(* IEC 61131-3 sources: plcassist-cli/packages/volt-lsp-iec/test-corpus/awa-palletizer/Device/Plc Logic/Application/Library Manager/L_TS2P_TechModulesSynchronizingCamming (part 2) *)

(* ---- L_TS2P_FLYINGSAWSTATE.fb ---- *)
FUNCTION_BLOCK L_TS2P_FLYINGSAWSTATE EXTENDS L_TB2P_TechModuleBase
VAR_INPUT
	XUSEORIGINAL : BOOL;
	XENABLE : BOOL;
	XENABLEOPERATION : BOOL;
	XRESETERROR : BOOL;
	XQSPAPPLICATION : BOOL;
	XABORT : BOOL;
	XJOGPOS : BOOL;
	XJOGNEG : BOOL;
	XHOMEEXECUTE : BOOL;
	LROVERRIDE : LREAL := 1;
	SCCTRLBASICMOTION : L_TB2P_scCtrlBasicMotion;
	SCPAR : L_TS2P_scPar_FlyingSawState;
	SCACCESSPOINTS : L_TS2P_scAP_FlyingSawState;
	MASTERVALUES : L_MC1P_IAXIS_REF_MASTERVALUES;
	XSTARTFLYINGSAW : BOOL;
	XSYNCININSTANT : BOOL;
	XEXECUTENEXTCUT : BOOL;
	XEXECUTEGAP : BOOL;
	XSETCUTTINGLENGTHINSTANT : BOOL;
	LRCUTTINGLENGTH : LREAL;
	LRSYNCOVERRIDE : LREAL := 1;
	XSETMATERIALCOUNTER : BOOL;
	XMOVETOPARKPOS : BOOL;
	XRESUMETARGETPOS : BOOL;
	XRESETMARKSTACK : BOOL;
	SCTPRECDATA_MARKSENSOR : L_MC1P.L_MC1P_TpReceiveData;
END_VAR
VAR_OUTPUT
	XREADYFOROPERATION : BOOL;
	XOPERATIONENABLED : BOOL;
	XREADYFORMOTION : BOOL;
	XERROR : BOOL;
	XWARNING : BOOL;
	EERRORID : L_IE1P_Error;
	XSTOACTIVE : BOOL;
	XQSPACTIVE : BOOL;
	XABORTBUSY : BOOL;
	XABORTDONE : BOOL;
	XJOGGINGBUSY : BOOL;
	XHOMINGBUSY : BOOL;
	XHOMINGDONE : BOOL;
	XISHOMED : BOOL;
	ETMSTATE : L_TB2P_States := L_TB2P_States.DISABLED;
	SCSTATUSBASICMOTION : L_TB2P_scStatusBasicMotion;
	LRACTVEL : LREAL;
	LRSETVELOUT : LREAL;
	LRACTPOS : LREAL;
	LRSETPOSOUT : LREAL;
	LRACTFOLLOWINGERROR : LREAL;
	SCSIGNALFLOW : L_TS2P_scSF_FlyingSawState;
	XSYNCHRONISED : BOOL;
	XACCDECSYNC : BOOL;
	XINPOSITION : BOOL;
	XPOSITIONING : BOOL;
	LRMATERIALCOUNTER : LREAL;
	LRTARGETPOS : LREAL;
	LRCUTGAP : LREAL;
	LRACTIVECUTTINGLENGTH : LREAL;
	WMARKSINSTACK : WORD;
END_VAR
VAR_IN_OUT
	AXIS : AXIS_REF;
END_VAR
VAR
	XINTERNALCONTROLACTIVE_OLD : BOOL;
	XUSEORIGINAL_OLD : BOOL;
	ITFCONNECTORFLYINGSAW : L_TS2P_IConnectorFlyingSaw;
	TM_INT : L_TS2M_TM_FlyingSawState;
	SCPAR_INT : L_TS2P_scPar_FlyingSawState;
	_SCDATA_INT : L_TS2M_scData_FlyingSawState;
	_SCFMDATA_INT : L_TS2M_scData_FM_FlyingSaw;
	_UICALLMFUNIDXINPUT : UINT := 1;
	_UICALLMFUNIDXOUTPUT : UINT := 1;
	_MCCALL : L_UM1P_MCCall;
	_ASCINPUT : ARRAY [1.._MCCall.c_BufferDepthInput] OF L_TS2P_FlyingSawStateIn;
	_ASCOUTPUT : ARRAY [1.._MCCall.c_BufferDepthOutput] OF L_TS2P_FlyingSawStateOut;
	_ASCPARCORE : ARRAY [1.._MCCall.c_BufferDepthInput] OF L_TS2P_scPar_FlyingSawState;
	_ASCACCESSPOINTSCORE : ARRAY [1.._MCCall.c_BufferDepthInput] OF L_TS2P_scAP_FlyingSawState;
	_ASCSIGNALFLOWCORE : ARRAY [1.._MCCall.c_BufferDepthOutput] OF L_TS2P_scSF_FlyingSawState;
	_ASCDATACORE : ARRAY [1.._MCCall.c_BufferDepthInput] OF L_TS2M_scData_FlyingSawState;
	_ASCDATAFMCORE : ARRAY [1.._MCCall.c_BufferDepthInput] OF L_TS2M_scData_FM_FlyingSaw;
	_SCINPUTVISU : L_TS2P_FlyingSawStateIn;
	_PSCINPUTVISU : POINTER TO L_TS2P_FlyingSawStateIn := ADR(_scInputVisu);
	_PSCOUTPUTVISU : POINTER TO L_TS2P_FlyingSawStateOut := ADR(_ascOutput[1]);
	_PSCPARVISU : POINTER TO L_TS2P_scPar_FlyingSawState := ADR(scPar_int);
	_PSCDATAVISU : POINTER TO L_TS2M_scData_FlyingSawState := ADR(_scData_int);
	_PSCFMDATAVISU : POINTER TO L_TS2M_scData_FM_FlyingSaw := ADR(_scFMData_int);
	_PSCFMSFVISU : POINTER TO L_TS2P_scSF_FlyingSawState;
	ITFBASICMOTIONBASE : L_TB2P.L_TB2P_IBasicMotionBase;
	ITFFLYINGSAWPROCESSINGEXTENSION : L_TS2P_IFlyingSawProcessing;
	ITFITECHMODULEINTERNAL : L_TB2P_ITechModuleInternal;
	LRJERKDEC : LREAL;
	LRJOGGINGJERKDEC : LREAL;
	REMAININGTIMEOFPROFILE : LREAL;
	REMAININGTIMEOFPROFILEAVAILABLE : BOOL;
END_VAR
END_FUNCTION_BLOCK

METHOD CALL_ABC
VAR_INPUT
	ITFTECHMODULE : L_TB2P.L_TB2P_IBasicMotionBase;
	XQSPAPPLICATION : BOOL;
	XHALT : BOOL;
	XABORT : BOOL;
	XHOMEEXECUTE : BOOL;
	XJOGPOS : BOOL;
	XJOGNEG : BOOL;
	XFINISHPOSITIONING : BOOL;
	XMOVEVELEXECUTE : BOOL;
	XMOVEABSEXECUTE : BOOL;
	XMOVERELEXECUTE : BOOL;
	XENABLEOPERATION : BOOL;
	XRESETERROR : BOOL;
	XENABLEPOSITIVE : BOOL;
	XENABLENEGATIVE : BOOL;
	XDISABLESWLIMIT : BOOL;
	LROVERRIDE : LREAL;
	LROVERRIDEACC : LREAL;
	LROVERRIDEJERK : LREAL;
	XRESETHOMEPOSITION : BOOL;
	XCONTINUOUSUPDATE : BOOL;
	LRPOS_DIST : LREAL;
	LRVEL : LREAL;
	LRACC : LREAL;
	LRDEC : LREAL;
	LRJERK : LREAL;
	EDIRECTION : L_TB2P.MC_DIRECTION;
	SCHOMEEXTTP : L_TB2P.MC_TRIGGER_REF;
	XHOMEABSSWITCH : BOOL;
	XSPECIALABORTBEHAVIOR : BOOL;
	LRABORTDEC : LREAL;
	LRABORTJERK : LREAL;
END_VAR
VAR_OUTPUT
	XERROR : BOOL;
	EERRORID : L_TB2P.L_IE1P_Error;
	XFUNBUSY : BOOL;
	XFUNDONE : BOOL;
	XFUNCOMMANDABORTED : BOOL;
	EFUNSTATEACT : L_TB2P.L_MC1P_ABC_State;
	ECONTROLMODE : L_TB2P.L_MC1P_ControlMode;
	XISHOMED : BOOL;
	XHWLIMITSWITCHNEG : BOOL;
	XHWLIMITSWITCHPOS : BOOL;
	XSWLIMITENABLED : BOOL;
	XSWLIMITSWITCHNEG : BOOL;
	XSWLIMITSWITCHPOS : BOOL;
	EAXISTYPE : L_TB2P.L_MC1P_DriveType;
	EAXISSTATE : L_TB2P.L_MC1P_AXIS_STATE;
	XSTOACTIVE : BOOL;
	XREADYFOROPERATION : BOOL;
	XOPERATIONENABLED : BOOL;
	XREADYFORMOTION : BOOL;
	XAXISWARNING : BOOL;
	XAXISERROR : BOOL;
	EAXISERRORID : L_TB2P.L_IE1P_Error;
	XDRIVEWARNING : BOOL;
	XDRIVEERROR : BOOL;
	DWDRIVEERRORID : DWORD;
	LRACTPOS : LREAL;
	LRACTVEL : LREAL;
	LRSETPOSOUT : LREAL;
	LRSETVELOUT : LREAL;
	LRACTFOLLOWINGERROR : LREAL;
	XINPOSITION : BOOL;
	XSTANDSTILLSETVELOCITY : BOOL;
	XSTANDSTILLACTVELOCITY : BOOL;
	XCONSTANTVELOCITY : BOOL;
	XACCELERATING : BOOL;
	XDECELERATING : BOOL;
	XDIRECTIONPOSITIVE : BOOL;
	XDIRECTIONNEGATIVE : BOOL;
	XAXISAVAILABLE : BOOL;
END_VAR
VAR_IN_OUT
	AXIS : AXIS_REF;
END_VAR
END_METHOD

METHOD GET_PAP : POINTER TO L_TB2P_scAP_TM_MotionControl
END_METHOD

METHOD GET_PDATA : POINTER TO L_TS2M_scData_FlyingSawState
END_METHOD

METHOD GET_PFMDATA : POINTER TO L_TS2M_scData_FM_FlyingSaw
END_METHOD

METHOD GET_PPAR : POINTER TO L_TB2P_scPar_TM_MotionControl
END_METHOD

METHOD GET_PSF : POINTER TO L_TB2P_scSF_TM_MotionControl
END_METHOD

METHOD CLUTCH
VAR_INPUT
	ITFTECHMODULE : L_TS2P_IFlyingSawProcessing;
	XENABLE : BOOL;
	XSYNCVEL : BOOL := FALSE;
	XSYNCPOS : BOOL;
	XSYNCOUTINSTANT : BOOL;
	LRSYNCVEL : LREAL := 10;
	LRSYNCACC : LREAL := 100;
	LRSYNCDEC : LREAL := 100;
	LRSYNCJERK : LREAL := 10000;
	LRCYCMASTERPOS : LREAL;
	LRCYCMASTERVEL : LREAL;
	LRCYCMASTERACC : LREAL;
	LRSETSLAVEPOS : LREAL;
	LRSETSLAVEVEL : LREAL;
	LRSETSLAVEACC : LREAL;
END_VAR
VAR_OUTPUT
	EERRORID : L_IE1P.L_IE1P_Error;
	XERROR : BOOL;
	XBUSY : BOOL;
	XDONE : BOOL;
	XACCDECSYNC : BOOL;
	XVELSYNCHRONISED : BOOL;
	XPOSSYNCHRONISED : BOOL;
	LRSETSLAVEPOSOUT : LREAL;
	LRSETSLAVEVELOUT : LREAL;
	LRSETSLAVEACCOUT : LREAL;
	XPROFILERESETTIMEVALID : BOOL;
	LRPROFILERESETTIME : LREAL;
END_VAR
END_METHOD

METHOD EXECUTEGAP
VAR_INPUT
	ITFTECHMODULE : L_TS2P_IFlyingSawProcessing;
	XENABLE : BOOL;
	LRSYNCVEL : LREAL := 10;
	LRSYNCACC : LREAL := 100;
	LRSYNCDEC : LREAL := 100;
	LRSYNCJERK : LREAL := 10000;
	XEXECUTEGAP : BOOL;
	XAUXEXECUTEGAP : BOOL := FALSE;
	LRCYCMASTERPOS : LREAL;
	LRCYCMASTERVEL : LREAL;
	LRCYCMASTERACC : LREAL;
	LRSETSLAVEPOS : LREAL;
	LRSETSLAVEVEL : LREAL;
	LRSETSLAVEACC : LREAL;
END_VAR
VAR_OUTPUT
	EERRORID : L_IE1P.L_IE1P_Error;
	XERROR : BOOL;
	XBUSY : BOOL;
	XDONE : BOOL;
	XACCDECSYNC : BOOL;
	XVELSYNCHRONISED : BOOL;
	XPOSSYNCHRONISED : BOOL;
	LRSETSLAVEPOSOUT : LREAL;
	LRSETSLAVEVELOUT : LREAL;
	LRSETSLAVEACCOUT : LREAL;
	XPROFILERESETTIMEVALID : BOOL;
	LRPROFILERESETTIME : LREAL;
END_VAR
END_METHOD

METHOD MARKSTACK_GETMARK
VAR_INPUT
	ITFTECHMODULE : L_TS2P_IFlyingSawProcessing;
	XENABLE : BOOL;
	XGETMARK : BOOL;
	XRESETGETMARK : BOOL;
	XRESETMARKSTACK : BOOL;
	LRCYCSETPOS : LREAL;
	LRCYCSETVEL : LREAL;
END_VAR
VAR_OUTPUT
	XMARKSTACKFULL : BOOL;
	XMARKSTACKEMPTY : BOOL;
	WMARKSINSTACK : WORD;
	XMARKVALID : BOOL;
	LRMARKPOSOUT : LREAL;
END_VAR
END_METHOD

METHOD MARKSTACK_SETMARK
VAR_INPUT
	ITFTECHMODULE : L_TS2P_IFlyingSawProcessing;
	XENABLE : BOOL;
	XSETMARK : BOOL;
	LRMARKPOS : LREAL;
	XRESETMARKSTACK : BOOL;
	LRCYCSETPOS : LREAL;
	LRCYCSETVEL : LREAL;
END_VAR
VAR_OUTPUT
	XMARKSTACKFULL : BOOL;
	XMARKSTACKEMPTY : BOOL;
	WMARKSINSTACK : WORD;
	XNEWMARKRECEIVED : BOOL;
END_VAR
END_METHOD

METHOD POSITIONING
VAR_INPUT
	ITFTECHMODULE : L_TS2P_IFlyingSawProcessing;
	XENABLE : BOOL;
	XMOVETOTARGETPOS : BOOL;
	LRTARGETPOS : LREAL;
	LRPOSITIONINGVEL : LREAL;
	LRPOSITIONINGACC : LREAL;
	LRPOSITIONINGDEC : LREAL;
	LRPOSITIONINGJERK : LREAL;
	LRSETSLAVEPOS : LREAL;
	LRSETSLAVEVEL : LREAL;
	LRSETSLAVEACC : LREAL;
	LRCORRECTTIMEBASE : LREAL := 0;
	LROVERRIDE : LREAL := 1.0;
END_VAR
VAR_OUTPUT
	EERRORID : L_IE1P.L_IE1P_Error;
	XERROR : BOOL;
	XBUSY : BOOL;
	XDONE : BOOL;
	XPOSITIONING : BOOL;
	XINPOSITION : BOOL;
	LRSETSLAVEPOSOUT : LREAL;
	LRSETSLAVEVELOUT : LREAL;
	LRSETSLAVEACCOUT : LREAL;
	XPROFILERESETTIMEVALID : BOOL;
	LRPROFILERESETTIME : LREAL;
END_VAR
END_METHOD

METHOD REQUESTINTERFACE : BOOL
VAR_INPUT
	ID : DINT;
	PITFUNKNOWN : POINTER TO L_UBUP.L_UBUP_IUnknown;
END_VAR
END_METHOD

METHOD CALLFUNCTION
VAR_INPUT
	UIINPUTDATAIDX : UINT;
	UIOUTPUTDATAIDX : UINT;
END_VAR
END_METHOD

METHOD COPYINPUTS : BOOL
VAR_INPUT
	IDX : WORD;
END_VAR
END_METHOD

METHOD COPYOUTPUTS : BOOL
VAR_INPUT
	IDX : WORD;
END_VAR
END_METHOD

METHOD FUNCTIONWASCALLEDTWICE : BOOL
VAR_INPUT
	IDX : WORD;
END_VAR
END_METHOD

METHOD HANDLESTANDARDCALL : BOOL
END_METHOD

METHOD SYNCOUTPUTS
VAR_INPUT
	UICOPYOUTPUTFROMIDX : UINT;
	UICOPYOUTPUTTOIDX : UINT;
END_VAR
END_METHOD

METHOD FB_INIT : BOOL
VAR_INPUT
	BINITRETAINS : BOOL;
	BINCOPYCODE : BOOL;
END_VAR
END_METHOD

METHOD CALL_INTERNALCTRL
END_METHOD

(* ---- L_TS2P_INVERTGEARFACTOR.fb ---- *)
FUNCTION_BLOCK L_TS2P_INVERTGEARFACTOR
VAR_INPUT
	XINVERTGEARFACTOR : BOOL;
	LRCYCLELENGTHX : LREAL := 1.0;
	LRCYCLELENGTHY : LREAL := 1.0;
	LRCOUPLINGX : LREAL := 1.0;
	LRCOUPLINGY : LREAL := 1.0;
	XDISABLETOLERANCEINVERTGEARFACTOR : BOOL;
	LRTOLERANCEINVERTGEARFACTOR : LREAL := 0;
END_VAR
VAR_OUTPUT
	XINVERTGEARFACTORACTIVE : BOOL;
	LRCYCLELENGTHX_OUT : LREAL;
	LRCYCLELENGTHY_OUT : LREAL;
	LRCOUPLINGX_OUT : LREAL;
	LRCOUPLINGY_OUT : LREAL;
	XWARNING : BOOL;
	EERRORID : L_IE1P_Error;
END_VAR
VAR_IN_OUT
	AXIS : AXIS_REF;
END_VAR
VAR
	XINWINDOW : BOOL;
END_VAR
END_FUNCTION_BLOCK

(* ---- L_TS2P_MARKQUEUE.fb ---- *)
FUNCTION_BLOCK L_TS2P_MARKQUEUE
VAR_INPUT
	XENABLE : BOOL;
	XLOADMARKPOS : BOOL;
	LRMARKPOS : LREAL;
	XGETNEXTMARK : BOOL;
	XRESETGETNEXTMARK : BOOL;
	XRESETMARKQUEUE : BOOL;
	LRCYCSETPOS : LREAL;
	LRCYCSETVEL : LREAL;
END_VAR
VAR_OUTPUT
	XQUEUEISFULL : BOOL;
	XQUEUEISEMPTY : BOOL;
	XNEWMARKRECEIVED : BOOL;
	WMARKSINQUEUE : WORD;
	XMARKVALID : BOOL;
	LRMARKPOSOUT : LREAL;
END_VAR
VAR
	FB_MB1P_STACK : L_MB1P_Stack;
	XTRACKMARK : BOOL;
	XENABLE_OLD : BOOL;
	XRESETMARKQUEUE_OLD : BOOL;
	XGETNEXTMARK_OLD : BOOL;
	XRESETGETNEXTMARK_OLD : BOOL;
	C_LRMATERIALCOUNTERCYCLELENGTH : LREAL := (16#4FFFFFFFFFFFFFFF * 1E-08);
END_VAR
END_FUNCTION_BLOCK

(* ---- L_TS2P_MARKSTACK.fb ---- *)
FUNCTION_BLOCK L_TS2P_MARKSTACK
VAR_INPUT
	XENABLE : BOOL;
	TPRECDATAIN : L_MC1P_TpReceiveData;
	LRACTVELMATERIAL : LREAL;
	LRACTPOSITIONTPAXIS : LREAL;
	LRCYCLELENGTHTPAXIS : LREAL;
	LRMARKSTACKLENGTH : LREAL;
	LRTASKCYCLE : LREAL;
END_VAR
VAR_OUTPUT
	TPRECDATAOUT : L_MC1P_TpReceiveData;
	XERROR : BOOL := FALSE;
	EERRORID : WORD;
	LRTPDIFFOUT : LREAL;
END_VAR
VAR
	ALRINTEGRATORSTARTPOS : ARRAY [1..64] OF LREAL := [64(0)];
	ALRLASTSCAN : ARRAY [1..64] OF LREAL := [64(0)];
	ALRDUMMY : ARRAY [1..64] OF LREAL := [64(0)];
	AXTPVALID : ARRAY [1..64] OF BOOL := [64(FALSE)];
	AXDUMMY : ARRAY [1..64] OF BOOL := [64(FALSE)];
	ADWACTTIMESTAMP : ARRAY [1..64] OF DWORD := [64(0)];
	ADWRECTIMESTAMP : ARRAY [1..64] OF DWORD := [64(0)];
	ADWDUMMY : ARRAY [1..64] OF DWORD := [64(0)];
	XREGISTERFULL : BOOL := FALSE;
	XINIT : BOOL := TRUE;
	WCOUNTER : WORD;
	WCOUNTERIN : WORD := 1;
	WCOUNTEROUT : WORD := 1;
	LRINTEGRATORPOS : LREAL := 0;
	LRCYCPOSDIFF : LREAL := 0;
	LRPOSTOREGISTEREND : LREAL := 0;
	XTPRECEIVEDINOLD : BOOL;
	LRMARKSTACKLENGTHOLD : LREAL;
	LRACTPOSITIONTPAXISCOMP : LREAL;
	LRACTTPPOSITIONOUT_INT : LREAL;
	DWDEADTIMESTACKOUT : DWORD;
	LRINTEGRATORLENGTH : LREAL := 10000000000.0;
END_VAR
END_FUNCTION_BLOCK

METHOD CALL_INITMARKSTACK
END_METHOD

(* ---- L_TS2P_MARKSTACKFLYINGSAW.fb ---- *)
FUNCTION_BLOCK L_TS2P_MARKSTACKFLYINGSAW
VAR
	FB_MB1P_STACK : L_MB1P_Stack_FlyingSaw;
	XTRACKMARK : BOOL;
	XMARKVALID_INT : BOOL;
	XENABLE_OLD : BOOL;
	XRESETMARKSTACK_OLD : BOOL;
	XGETMARK_OLD : BOOL;
	XSETMARK_OLD : BOOL;
	XRESETGETMARK_OLD : BOOL;
	C_LRMATERIALCOUNTERCYCLELENGTH : LREAL := (16#4FFFFFFFFFFFFFFF * 1E-08);
END_VAR
END_FUNCTION_BLOCK

METHOD DISABLE
END_METHOD

METHOD RESETMARKSTACK
END_METHOD

METHOD GETMARK
VAR_INPUT
	XENABLE : BOOL;
	XGETMARK : BOOL;
	XRESETGETMARK : BOOL;
	XRESETMARKSTACK : BOOL;
	LRCYCSETPOS : LREAL;
	LRCYCSETVEL : LREAL;
END_VAR
VAR_OUTPUT
	XMARKSTACKFULL : BOOL;
	XMARKSTACKEMPTY : BOOL;
	WMARKSINSTACK : WORD;
	XMARKVALID : BOOL;
	LRMARKPOSOUT : LREAL;
END_VAR
END_METHOD

METHOD SETMARK
VAR_INPUT
	XENABLE : BOOL;
	XSETMARK : BOOL;
	LRMARKPOS : LREAL;
	XRESETMARKSTACK : BOOL;
	LRCYCSETPOS : LREAL;
	LRCYCSETVEL : LREAL;
END_VAR
VAR_OUTPUT
	XMARKSTACKFULL : BOOL;
	XMARKSTACKEMPTY : BOOL;
	WMARKSINSTACK : WORD;
	XNEWMARKRECEIVED : BOOL;
END_VAR
END_METHOD

(* ---- L_TS2P_MARKWINDOWRELATIVE.fb ---- *)
FUNCTION_BLOCK L_TS2P_MARKWINDOWRELATIVE
VAR_INPUT
	XENABLE : BOOL;
	LRTPWINDOWSIZE : LREAL;
	LRSETOFFSETTPWINDOW : LREAL;
	LRCYCVEL : LREAL;
	TPRECDATAIN : L_MC1P_TpReceiveData;
	LRSTARTPOSITION : LREAL;
	LRCYCLELENGTH : LREAL;
	XTEACHMARKWINDOW : BOOL;
	DWMAXTPNOTDETECTED : DWORD;
	LRTASKCYCLE : LREAL;
END_VAR
VAR_OUTPUT
	TPRECDATAOUT : L_MC1P_TpReceiveData;
	XTPWINDOWOPEN : BOOL;
	XTPWINDOWOPENCOMP : BOOL;
	LRTPDELTAPOSCOMP : LREAL;
	XTPINWINDOW : BOOL;
	XTPNOTINWINDOW : BOOL;
	XTPNOTDETECTED : BOOL;
	XTPSENSORTEACHED : BOOL;
	XMAXTPNOTDETECTED : BOOL;
END_VAR
VAR
	LRMARKWINDOWINTEGRATOROLD : LREAL;
	XTPNOTDETECTEDINTERNAL : BOOL;
	LRLOWERWINDOW : LREAL;
	LRUPPERWINDOW : LREAL;
	XTEACHTPSENSOROLD : BOOL;
	DWMISSEDTPCOUNTER : DWORD;
	XTPISINWINDOW : BOOL;
	LRDEADTIMEPOSDIFF : LREAL;
	LRUPPERWINDOWCOMP : LREAL;
	XTPCOMPWINDOWOPEN : BOOL;
	XTPCOMPWINDOWOPENOLD : BOOL := FALSE;
	LRLOWERWINDOWCOMP : LREAL;
	XTPRECEIVEDOLD : BOOL;
	XTPRECEIVEDINTERNAL : BOOL;
	LRTPWINDOWSIZE_INT : LREAL;
	LRMARKWINDOWINTEGRATOR : LREAL := 0;
	LRDEADTIMETP : LREAL;
	LRACTUALTPPOSITION : LREAL;
END_VAR
END_FUNCTION_BLOCK

(* ---- L_TS2P_MASTERVALUECORRECTION.fb ---- *)
FUNCTION_BLOCK L_TS2P_MASTERVALUECORRECTION
VAR_INPUT
	XAXIS : POINTER TO L_MC1P_IAXIS_REF_MASTERVALUES;
	XENABLE : BOOL;
	XENABLECORRECTION : BOOL;
	XRESETERROR : BOOL;
	LRSETVELIN : LREAL;
	LRACTPOSITIONTOOL : LREAL;
	LRCYCLELENGTHTOOL : LREAL;
	TPRECDATA : L_MC1P_TpReceiveData;
	XLOADREGPOS : BOOL;
	LRLOADREGPOS : LREAL;
	LRSENSORTOOLDIST : LREAL;
	LRMARKDIST : LREAL;
	LRMAXCORRNEG : LREAL;
	LRMAXCORRPOS : LREAL;
	ESOURCEFORCORRWINDOW : L_TS2P_SourceForCorrWindow;
	LRUPPERCORRPOS : LREAL;
	LRLOWERCORRPOS : LREAL;
	DWGEARINGNUMERATORY : DWORD := 1;
	DWGEARINGDENOMINATORY : DWORD := 1;
	XSYNCHRONISED : BOOL;
	LRACTOFFSETMASTERIN : LREAL;
	LRACTOFFSETSLAVEIN : LREAL;
	XTEACHMARKWINDOW : BOOL;
	XENABLEMARKWINDOW : BOOL;
	LRMARKWINDOWSIZE : LREAL;
	LRSETOFFSETMARKWINDOW : LREAL;
	DWMAXNUMBERVIRTUALMARKS : DWORD;
	LRGEARFACTORCORRGAIN : LREAL;
	LRMAXGEARFACTORCORR : LREAL;
	XGEARFACTORCORR : BOOL;
	XGEARFACTORCORRHOLD : BOOL;
	XENABLETOOLCORRECTION : BOOL;
	LRTRANSMITCYCLESSETPOS : LREAL;
	DIDEADTIMECOMP : DINT;
	LRCORRVEL : LREAL;
	LRCORRACC : LREAL;
	LRCORRDEC : LREAL;
	LRCORRJERK : LREAL;
	ECORRMODE : L_TS2P_CorrectionMode;
	ECORRMODEOLD : L_TS2P_CorrectionMode;
END_VAR
VAR_OUTPUT
	CORRECTEDXAXIS : L_MC1P_IAXIS_REF_MASTERVALUES;
	LRACTVEL : LREAL;
	XERROR : BOOL;
	XWARNING : BOOL;
	EERRORID : WORD;
	XCORRLIMITED : BOOL;
	LRACTMARKERROR : LREAL;
	LRACTMARKDIST : LREAL;
	XINITDONE : BOOL;
	XCORRACTIVE : BOOL;
	XMARKRECEIVED : BOOL;
	LRSENSORACTPOS : LREAL;
	LRSENSORSETPOS : LREAL;
	XMARKWINDOWOPEN : BOOL;
	XMARKOUTOFWINDOW : BOOL;
	XMARKNOTDETECTED : BOOL;
	XMARKWINDOWTEACHED : BOOL;
	LRGEARFACTORCORR : LREAL;
	XGEARFACTORCORRLIMITED : BOOL;
	XCORRNEXTCYCLE : BOOL;
END_VAR
VAR_IN_OUT
	YAXIS : AXIS_REF;
END_VAR
VAR
	FB_L_TB2P_TP_CONVERTER : L_TB2P_TP_Converter;
	FB_L_TS2P_MARKWINDOWRELATIVE : L_TS2P_MarkWindowRelative;
	FB_L_TS2P_TPVIRTUALACTPOS : L_TS2P_TpVirtualActPos;
	FB_L_TS2P_MARKSTACK : L_TS2P_MarkStack;
	FB_L_MC1P_TPCALCDIFF : L_MC1P_TpCalcDiff;
	FB_L_TS2P_TPLIMITDIFF : L_TS2P_TpLimitDiff;
	FB_L_TS2P_DISTCORRECTIONWINDOW : L_TS2P_DistCorrectionWindow;
	FB_L_MC1P_SETAXISREFMASTERVALUES : L_MC1P_SetAxisRefMasterValues;
	FB_PROFILEGENERATOR : L_MC1P_ProfileGenerator;
	FB_INTEGRATOR : L_MC1P_IntegrateAxis;
	SCPROFILEPARAMETER : L_MC1P_ProfileParameter;
	FB_RAMPGENERATORGEARFACTOR : L_MC1P_RampGenerator;
	LRSENSORSETPOS_INT : LREAL;
	LRGEARINGFAKTOR : LREAL := 1.0;
	LRTPDIFFERENCE_INT : LREAL;
	XTPINWINDOW : BOOL;
	XVALUESTOREDTPCONVERTER : BOOL;
	XVALUESTOREDTPCONVERTEROLD : BOOL;
	XVALUESTOREDMARKWINDOW : BOOL;
	XVALUESTOREDMISSEDMARKS : BOOL;
	XVALUESTOREDMARKSTACK : BOOL;
	XVALUESTOREDCALCDIFF : BOOL;
	XVALUESTOREDLIMIT : BOOL;
	LRCORRRESIDUAL : LREAL;
	LRTPACTPOSITION_INT : LREAL;
	LRTPDIFFERENCELIM_INT : LREAL;
	LROFFSETPOSCTRL_INT : LREAL;
	LRCYCVELIN_INT : LREAL;
	LRSETCORRECTEDPOSOUT_INT : LREAL;
	LRMASTERSETPOSOLD_INT : LREAL;
	LRCORRPOSOUTOLD_INT : LREAL;
	LRVELOUT_INT : LREAL;
	XCORRACTIVE_INT : BOOL;
	XINIT : BOOL := TRUE;
	XTPCORRECTIONACTIVE : BOOL := FALSE;
	LRTPAXISSETPOS : LREAL;
	LRMARKDIST_INT : LREAL;
	XZERO : BOOL;
	XHOMINGDONE : BOOL;
	XSTARTREFERENCEACTIVE : BOOL;
	XHOMINGACTIVE : BOOL := FALSE;
	XMARKDISTCHANGED : BOOL;
	XENABLE_OLD : BOOL;
	XTPRECEIVEDOUT_INTOLD : BOOL;
	XSTARTFIRSTCORRECTION : BOOL;
	LRTPDIFFERENCELIM2_INT : LREAL;
	XCORRECTIONBUSYOLD : BOOL;
	LRTPACTPOSIN_OLD : LREAL;
	LRTPSETPOSIN_OLD : LREAL;
	LRTPAXISACTPOS_OLD : LREAL;
	LRCYCLELENGTH : LREAL;
	ICOUNTER : INT := 0;
	LRSETPOSITIONOLD : LREAL;
	LRCYCLELENGTHTP : LREAL;
	LRTPACTPOSITIONOLD : LREAL;
	XFIRSTTOUCHPROBE : BOOL := TRUE;
	LRSENSORTOOLDISTANCE_INT : LREAL;
	LRMARKSTACKLENGTH : LREAL;
	LRTPDIFFERENCELIMITOUT_INT : LREAL;
	XTPNOTDETECTED_INT : BOOL;
	XMAXTPNOTDETECTED : BOOL;
	LRGEARINGFAKTOROLD : LREAL;
	LRGEARFACTORINTEGRATOR : LREAL;
	LRGEARFACTORGAIN : LREAL := 1;
	LRGEARFACTORNUMERATORCORR : LREAL;
	LRGEARFACTORNUMERATORCORRLIMITED : LREAL;
	LRGEARFACTORDENOMINATOR : LREAL;
	LRGEARFACTORNUMERATOR : LREAL;
	LRTOTALSTACKDIFFERENCEOUT_INT : LREAL := 0;
	LCORRECTIONVELIN : LREAL;
	LRSETPOSCORROUT_OLD : LREAL;
	LRDELTAGEARFACTORCORR : LREAL;
	XTPSENSORTEACHEDOLD : BOOL;
	XTPSENSORTEACHEDATLASTMARK : BOOL;
	XCALCMARKDISTINITIALISED : BOOL;
	XTEACHTPSENSOROLD : BOOL;
	LRTPDEADTIMEDIFF : LREAL;
	XTPRECEIVEDOUTOLD_INT : BOOL;
	LRMARKDISTINTEGRATOR : LREAL;
	LRTPAXISCOMPFACTOR : LREAL;
	LRTPAXISDELAYCYCLE : LREAL;
	XENABLEOLD : BOOL;
	XTPRECEIVEDINOLD_INT : BOOL;
	TPRECDATAMARKWINDOW : L_MC1P_TpReceiveData;
	TPRECDATAMARKSTACK : L_MC1P_TpReceiveData;
	LRMASTERACTPOSITIONOLD_INT : LREAL;
	XFIRSTVALUESTORED : BOOL := FALSE;
	LRSETINTEGRATEDPOSITIONOLD : LREAL;
	XRESETERROROLD : BOOL;
	LRTPDIFF : LREAL;
	LRVELDIFF : LREAL;
	LRVELCOMP : LREAL;
	SETPOSITIONFORSYNCOLD : LREAL;
	LRMARKDISTOLD : LREAL;
END_VAR
END_FUNCTION_BLOCK

METHOD CALL_CALCACTMARKDIST
END_METHOD

METHOD CALL_CALCMARKERROR
END_METHOD

METHOD CALL_CORRECTIONPOS
END_METHOD

METHOD CALL_CORRECTIONPROFILE
END_METHOD

METHOD CALL_ENABLEREGISTERCONTROL
END_METHOD

METHOD CALL_ERRORHANDLER
END_METHOD

METHOD CALL_FB
VAR_IN_OUT
	YAXIS : AXIS_REF;
END_VAR
END_METHOD

METHOD CALL_GEARFACTORCORRECTION
END_METHOD

METHOD CALL_GEARING
END_METHOD

METHOD CALL_INPUT
END_METHOD

METHOD CALL_LIMIT
END_METHOD

METHOD CALL_MARKDISTCHANGE
END_METHOD

METHOD CALL_MARKSENSORPOS
END_METHOD

METHOD CALL_MARKSTACK
END_METHOD

METHOD CALL_MARKWINDOW
VAR_IN_OUT
	YAXIS : AXIS_REF;
END_VAR
END_METHOD

METHOD CALL_NOTENABLE
END_METHOD

METHOD CALL_OUTPUT
END_METHOD

METHOD CALL_RESET
END_METHOD

METHOD CALL_RESETOUTPUTS
END_METHOD

METHOD CALL_SETAXISREFMASTERVALUES
END_METHOD

METHOD CALL_TPCONVERTER
END_METHOD

METHOD CALL_VIRTUALACTPOS
END_METHOD

METHOD GET_ACTMARKERRORLIMITED : LREAL
END_METHOD

METHOD GET_ACTUALMARKDIST : LREAL
END_METHOD

METHOD GET_CORRREGPOS : LREAL
END_METHOD

METHOD GET_INTEGRATORREGPOS : LREAL
END_METHOD

METHOD GET_MARKERRORUNLIMITED : LREAL
END_METHOD

METHOD GET_MARKPOSITIONINREGISTER : LREAL
END_METHOD

METHOD GET_MARKRECEIVEUNLIMITED : BOOL
END_METHOD

METHOD GET_MARKRECEIVEDLIMITED : BOOL
END_METHOD

METHOD GET_MARKWINDOWCOMP : BOOL
END_METHOD

METHOD GET_REGISTERINPUTVEL : LREAL
END_METHOD

METHOD GET_SETVELOCITYREGISTER : LREAL
END_METHOD

METHOD GET_LRMARKSTACKLENGTH : LREAL
END_METHOD

METHOD SETTPCOMPFACTOR : LREAL
END_METHOD

METHOD SETTPDELAYCYCLE : LREAL
END_METHOD

(* ---- L_TS2P_MATERIALCOUNTER.fb ---- *)
FUNCTION_BLOCK L_TS2P_MATERIALCOUNTER
VAR_INPUT
	XENABLE : BOOL;
	LRPOSIN : LREAL;
	LRTASKCYCLE : LREAL;
	LRPOSINSLAVE : LREAL;
	LRCYCLELEN : LREAL;
	XLOADSTARTPOS : BOOL;
	XSETMATERIALCOUNTER : BOOL;
	LRSETMATERIALPOS : LREAL;
	XLOADDELTAPOS : BOOL;
	LRSETDELTAPOS : LREAL;
	XSTARTFLYINGSAW : BOOL;
END_VAR
VAR_OUTPUT
	LNMATERIALPOS_E8 : LINT;
	LRMATERIALCOUNTER : LREAL;
	LRDELTAMATERIALPOS : LREAL;
END_VAR
VAR_IN_OUT
	AXIS : AXIS_REF;
END_VAR
VAR
	LNMODULOPOS_E8 : LINT;
	LNMODULOPOSOLD_E8 : LINT;
	LNCYCLELEN_E8 : LINT;
	LNPOSXDIFF : LINT;
	LNMATERIALPOS_E8_OLD : LINT;
	LNDELTAMATERIALPOS : LINT;
	XSETMATERIALCOUNTER_OLD : BOOL;
	XENABLE_OLD : BOOL;
END_VAR
END_FUNCTION_BLOCK

(* ---- L_TS2P_MULTICAMSEQUENCER.fb ---- *)
FUNCTION_BLOCK L_TS2P_MULTICAMSEQUENCER
VAR_INPUT
	XENABLE : BOOL;
	XCAMSEQUENCER : BOOL;
	EMODE : L_TS2P_CamSequenceMode;
	XCAMCHANGEINSTANT : BOOL;
	XLOADCAMTABLE : BOOL;
	WSETCAMTABLE : WORD;
	XENDOFPROFILEIN : BOOL;
	CAMTABLE1 : MC_CAM_REF;
	CAMTABLE2 : MC_CAM_REF;
	CAMTABLE3 : MC_CAM_REF;
	CAMTABLE4 : MC_CAM_REF;
END_VAR
VAR_OUTPUT
	XDONE : BOOL;
	XBUSY : BOOL;
	XERROR : BOOL;
	EERRORID : L_IE1P_Error;
	WACTIVECAMTABLE : WORD;
	CAMTABLEOUT : MC_CAM_REF;
	XCAMTABLEVALID : BOOL;
END_VAR
VAR
	WFMSTATE : WORD := 0;
	XINITSTATE : BOOL;
	XENABLE_OLD : BOOL;
	XLOADCAMTABLE_OLD : BOOL;
	XENDOFPROFILEIN_OLD : BOOL;
	XCAMSEQUENCER_OLD : BOOL;
	XCAMCHANGEINSTANT_OLD : BOOL;
	XCAMSEQUENCERACTIVE : BOOL;
END_VAR
END_FUNCTION_BLOCK

METHOD CALL_ERRORHANDLER
END_METHOD

METHOD CALL_FBMETHODS
END_METHOD

METHOD CALL_OUTPUT
END_METHOD

METHOD CALL_RESETCOMMANDS
END_METHOD

METHOD CALL_RESETOUTPUT
END_METHOD

METHOD CALL_STATEMACHINE
END_METHOD

METHOD CALL_SETCAMTABLEOUT
VAR_INPUT
	WSETCAMTABLE : WORD;
END_VAR
END_METHOD

METHOD CAMREFCHANGED : BOOL
VAR_IN_OUT
	CAMREFNEW : MC_CAM_REF;
	CAMREFOLD : MC_CAM_REF;
END_VAR
END_METHOD

METHOD SET_INIT
END_METHOD

METHOD CALL_S000_CYCLIC
END_METHOD

METHOD CALL_S001_INIT
END_METHOD

METHOD CALL_S002_READY
END_METHOD

METHOD CALL_S151_SEQUENCE_CYCLICCAM1
END_METHOD

METHOD CALL_S152_SEQUENCE_CYCLICCAM3
END_METHOD

METHOD CALL_S153_SEQUENCE_CAM1CYCLICCAM3CAM1
END_METHOD

METHOD CALL_S154_SEQUENCE_CAM1CAM2CYCLICCAM3CAM4CAM1
END_METHOD

(* ---- L_TS2P_OFFSETANDTRIM.fb ---- *)
FUNCTION_BLOCK L_TS2P_OFFSETANDTRIM
VAR_INPUT
	XENABLE : BOOL;
	LRSETOFFSET : LREAL;
	XLOADOFFSET : BOOL;
	XTRIMVELOCITY : BOOL;
	XTRIMPOS : BOOL;
	XTRIMNEG : BOOL;
	XRESETTRIMOFFSET : BOOL;
	EALLOWEDDIRECTION : L_TB2P_AllowedDirection;
	EACTDIRECTION : MC_DIRECTION;
	LRSETTRIMDISTANCE : LREAL;
	LRSETOFFSETTRIMVEL : LREAL := 100.0;
	LRSETOFFSETTRIMACC : LREAL := 1000.0;
	LRSETOFFSETTRIMDEC : LREAL := 1000.0;
	LRSETOFFSETTRIMJERK : LREAL := 100000.0;
	LRCYCMASTERPOS : LREAL;
	LRCYCMASTERVEL : LREAL;
	LRCYCMASTERACC : LREAL;
END_VAR
VAR_OUTPUT
	XBUSY : BOOL;
	XDONE : BOOL;
	XERROR : BOOL;
	EERRORID : WORD;
	LRSETOFFSETOUTTOTAL : LREAL;
	LRSETOFFSETOUT : LREAL;
	LRSETOFFSETOUTTRIM : LREAL;
	LRSETOFFSETOUTTOTALVEL : LREAL;
END_VAR
VAR
	XTRIMPOSOLD : BOOL := FALSE;
	XTRIMNEGOLD : BOOL := FALSE;
	XRESETTRIMOFFSETOLD : BOOL := FALSE;
	LRTRIMPOSITION : LREAL;
	XTRIMPOSEDGE : BOOL;
	XTRIMNEGEDGE : BOOL;
	XABORTPROFILEGENERATORTRIM : BOOL;
	LRTRIMDECDIST : LREAL;
	LRSETOFFSETTRIM_INT : LREAL;
	LRTARGETPOSOLD : LREAL;
	LRSETOFFSETTOTAL : LREAL;
	XPROFILEGENERATORACTIVEOFFSET : BOOL := FALSE;
	LRSETOFFSETOLD : LREAL;
	LRSETOFFSET_INT : LREAL;
	LRSETOFFSETOUTTOTALSAVE : LREAL;
	LRSETOFFSETSAVE : LREAL;
	LRSETPOSOUT_INT : LREAL;
	LRSETVELOUT_INT : LREAL;
	LRSETACCOUT_INT : LREAL;
	LRSETOFFSETTRIMVEL_INT : LREAL;
	LRSETOFFSETTRIMACC_INT : LREAL;
	LRSETOFFSETTRIMDEC_INT : LREAL;
	LRSETOFFSETTRIMJERK_INT : LREAL;
	LRSETOFFSETTRIMVELOLD_INT : LREAL;
	LRSETOFFSETTRIMACCOLD_INT : LREAL;
	LRSETOFFSETTRIMDECOLD_INT : LREAL;
	LRSETOFFSETTRIMJERKOLD_INT : LREAL;
	XMASTERVELDISABLEDDIRECTION : BOOL := FALSE;
	XMASTERVELDISABLEDDIRECTIONOLD : BOOL;
	XEXECUTEPOSITIONING : BOOL;
	XABORTPOSITIONING : BOOL;
	XAUXEXECUTE : BOOL;
	XABORTPOSITIVE : BOOL;
	XINITDONE : BOOL := FALSE;
	LRTASKCYCLETIME : LREAL := 0.001;
	XLOADOFFSET_OLD : BOOL;
	PROFILEGENERATOR : L_MC1P_ProfileGenerator;
	SCPROFILEPARAMETER : L_MC1P_ProfileParameter;
	LRSETOFFSETOUTTOTAL_OLD : LREAL;
END_VAR
END_FUNCTION_BLOCK

METHOD CALL_ADDOFFSETS
END_METHOD

METHOD CALL_AVOIDREVERSING
END_METHOD

METHOD CALL_INITROUTINE
END_METHOD

METHOD CALL_INPUTS
END_METHOD

METHOD CALL_LOADOFFSET
END_METHOD

METHOD CALL_OUTPUT
END_METHOD

METHOD CALL_PROFILEGENERATOR
END_METHOD

METHOD CALL_RESETOUTPUT
END_METHOD

METHOD CALL_TRIMING
END_METHOD

(* ---- L_TS2P_PROCESSCONTROL.fb ---- *)
FUNCTION_BLOCK L_TS2P_PROCESSCONTROL
VAR_INPUT
	XENABLE : BOOL;
	XSYNCFLYINGSAW : BOOL;
	XSYNCININSTANT : BOOL;
	XEXECUTEFIRSTCUT : BOOL;
	XRESUMETARGETPOS : BOOL;
	XRESET : BOOL;
	XTPNOTVALID : BOOL;
	XEXECUTEGAP : BOOL;
	XSETCUTTINGLENGTHINSTANT : BOOL;
	XDONEPROFILE : BOOL;
	LRSLAVEPOSIN : LREAL;
	LRLOWERLIMIT : LREAL;
	LRUPPERLIMIT : LREAL;
	LRSTARTPOS : LREAL;
	LRPOSX1 : LREAL;
	LRVELX1 : LREAL;
	LRACCX1 : LREAL;
	LRTASKCYCLE : LREAL;
END_VAR
VAR_OUTPUT
	XEXECUTEPROFILE : BOOL;
	XAUXEXECUTEPROFILE : BOOL;
	XSYNCPOSOUT : BOOL;
	LRPOSX2 : LREAL;
	LRVELX2 : LREAL;
	LRACCX2 : LREAL;
	XCUTTINGACTIVE : BOOL;
	LRTOLERANCE : LREAL;
	XTARGETOUTSIDELOWERLIMIT : BOOL;
	LRRESTTIMETARGETTOLOWERLIMIT : LREAL;
	LRDISTTOTARGET : LREAL;
END_VAR
VAR
	XEXECUTEPROFILE_INT : BOOL;
	XSYNC_INT : BOOL;
	WSTEPPER : WORD;
	XEXECUTEGAP_OLD : BOOL;
	XRESET_OLD : BOOL;
	XSYNCININSTANT_OLD : BOOL;
	XENABLE_OLD : BOOL;
	LRSTARTTHRESHOLD : LREAL;
	XSETCUTTINGLENGTHINSTANT_OLD : BOOL;
	XRESUMETARGETPOS_OLD : BOOL;
	XEXECUTEFIRSTCUT_OLD : BOOL;
	XMATERIALCONSTANTVEL : BOOL;
	LRMATERIALVEL : LREAL;
	LRMATERIALACC : LREAL;
	XSYNCININSTANT_LOCK : BOOL;
END_VAR
END_FUNCTION_BLOCK

(* ---- L_TS2P_SYNCANDCORRECTIONSTATE.fb ---- *)
FUNCTION_BLOCK L_TS2P_SYNCANDCORRECTIONSTATE EXTENDS L_TB2P_TechModuleBase
VAR_INPUT
	XUSEORIGINAL : BOOL;
	XENABLE : BOOL;
	XENABLEOPERATION : BOOL;
	XRESETERROR : BOOL;
	XQSPAPPLICATION : BOOL;
	XABORT : BOOL;
	XJOGPOS : BOOL;
	XJOGNEG : BOOL;
	XHOMEEXECUTE : BOOL;
	LROVERRIDE : LREAL := 1;
	SCCTRLBASICMOTION : L_TB2P_scCtrlBasicMotion;
	SCPAR : L_TS2P_scPar_SyncAndCorrectionState;
	SCACCESSPOINTS : L_TS2P_scAP_SyncAndCorrectionState;
	MASTERVALUES : L_MC1P_IAXIS_REF_MASTERVALUES;
	XSYNCIN : BOOL;
	XSYNCPOSRESTORE : BOOL;
	LRSETBASEVEL : LREAL;
	LRSETOFFSETPOS : LREAL;
	XTRIMPOS : BOOL;
	XTRIMNEG : BOOL;
	XTRIMRESET : BOOL;
	SCTPRECDATA_MARKSENSOR : L_MC1P_TpReceiveData;
	SCTPRECDATA_TOOLSENSOR : L_MC1P_TpReceiveData;
	XTEACHMARKWINDOW : BOOL;
	XTEACHMARKWINDOWTOOL : BOOL;
	XGEARFACTORCORR : BOOL;
	XGEARFACTORCORRHOLD : BOOL;
END_VAR
VAR_OUTPUT
	XREADYFOROPERATION : BOOL;
	XOPERATIONENABLED : BOOL;
	XREADYFORMOTION : BOOL;
	XERROR : BOOL;
	XWARNING : BOOL;
	EERRORID : L_IE1P_Error;
	XSTOACTIVE : BOOL;
	XQSPACTIVE : BOOL;
	XABORTBUSY : BOOL;
	XABORTDONE : BOOL;
	XJOGGINGBUSY : BOOL;
	XHOMINGBUSY : BOOL;
	XHOMINGDONE : BOOL;
	XISHOMED : BOOL;
	ETMSTATE : L_TB2P_States := L_TB2P_States.DISABLED;
	SCSTATUSBASICMOTION : L_TB2P_scStatusBasicMotion;
	LRACTVEL : LREAL;
	LRSETVELOUT : LREAL;
	LRACTPOS : LREAL;
	LRSETPOSOUT : LREAL;
	LRACTFOLLOWINGERROR : LREAL;
	SCSIGNALFLOW : L_TS2P_scSF_SyncAndCorrectionState;
	XSYNCHRONISED : BOOL;
	XACCDECSYNC : BOOL;
	XOFFSETTRIMACTIVE : BOOL;
	XBASEVELOCITYACTIVE : BOOL;
	LROFFSETTOTAL : LREAL;
	LRSETMARKCORROUT : LREAL;
	XMARKWINDOWTEACHED : BOOL;
	LRGEARFACTORCORR : LREAL;
	LRSETTOOLCORROUT : LREAL;
	XMARKWINDOWTEACHEDTOOL : BOOL;
END_VAR
VAR_IN_OUT
	AXIS : AXIS_REF;
END_VAR
VAR
	XINTERNALCONTROLACTIVE_OLD : BOOL;
	ITFCONNECTORSYNCANDCORRECTION : L_TS2P_IConnectorSyncAndCorrection;
	TM_INT : L_TS2P_TM_SyncAndCorrectionState;
	SCPAR_INT : L_TS2P_scPar_SyncAndCorrectionState;
	SCDATA_INT : L_TS2P_scData_TM_SyncAndCorrectionState;
	SCDATASP_INT : L_TS2P_scData_TM_SyncPosBase;
	XUSEORIGINAL_OLD : BOOL;
	_UICALLMFUNIDXINPUT : UINT := 1;
	_UICALLMFUNIDXOUTPUT : UINT := 1;
	_MCCALL : L_UM1P_MCCall;
	_ASCINPUT : ARRAY [1.._MCCall.c_BufferDepthInput] OF L_TS2P_SyncAndCorrectionStateIn;
	_ASCOUTPUT : ARRAY [1.._MCCall.c_BufferDepthOutput] OF L_TS2P_SyncAndCorrectionStateOut;
	_ASCPARCORE : ARRAY [1.._MCCall.c_BufferDepthInput] OF L_TS2P_scPar_SyncAndCorrectionState;
	_ASCACCESSPOINTSCORE : ARRAY [1.._MCCall.c_BufferDepthInput] OF L_TS2P_scAP_SyncAndCorrectionState;
	_ASCSIGNALFLOWCORE : ARRAY [1.._MCCall.c_BufferDepthOutput] OF L_TS2P_scSF_SyncAndCorrectionState;
	_SCINPUTVISU : L_TS2P_SyncAndCorrectionStateIn;
	_PSCINPUTVISU : POINTER TO L_TS2P_SyncAndCorrectionStateIn := ADR(_scInputVisu);
	_PSCOUTPUTVISU : POINTER TO L_TS2P_SyncAndCorrectionStateOut := ADR(_ascOutput[1]);
	_PSCDATAVISU : POINTER TO L_TS2P_scData_TM_SyncAndCorrectionState := ADR(scData_int);
	_PSCDATASPVISU : POINTER TO L_TS2P_scData_TM_SyncPosBase := ADR(scDataSP_int);
	_PSCPARVISU : POINTER TO L_TS2P_scPar_SyncAndCorrectionState := ADR(scPar_int);
	_PSCAPVISU : POINTER TO L_TS2P_scAP_SyncAndCorrectionState;
	_PSCSFVISU : POINTER TO L_TS2P_scSF_SyncAndCorrectionState;
	ITFBASICMOTIONBASE : L_TB2P.L_TB2P_IBasicMotionBase;
	ITFITECHMODULEINTERNAL : L_TB2P_ITechModuleInternal;
	ITFSYNCANDCORRECTIONEXTENSION : L_TS2P_ISyncAndCorrectionState;
	ITFSYNCPOSEXTENSION : L_TS2P_ISyncPosBase;
	LRJERKDEC : LREAL;
	LRJOGGINGJERKDEC : LREAL;
	REMAININGTIMEOFPROFILE : LREAL;
	REMAININGTIMEOFPROFILEAVAILABLE : BOOL;
END_VAR
END_FUNCTION_BLOCK

METHOD CALL_ABC
VAR_INPUT
	ITFTECHMODULE : L_TB2P.L_TB2P_IBasicMotionBase;
	XQSPAPPLICATION : BOOL;
	XHALT : BOOL;
	XABORT : BOOL;
	XHOMEEXECUTE : BOOL;
	XJOGPOS : BOOL;
	XJOGNEG : BOOL;
	XFINISHPOSITIONING : BOOL;
	XMOVEVELEXECUTE : BOOL;
	XMOVEABSEXECUTE : BOOL;
	XMOVERELEXECUTE : BOOL;
	XENABLEOPERATION : BOOL;
	XRESETERROR : BOOL;
	XENABLEPOSITIVE : BOOL;
	XENABLENEGATIVE : BOOL;
	XDISABLESWLIMIT : BOOL;
	LROVERRIDE : LREAL;
	LROVERRIDEACC : LREAL;
	LROVERRIDEJERK : LREAL;
	XRESETHOMEPOSITION : BOOL;
	XCONTINUOUSUPDATE : BOOL;
	LRPOS_DIST : LREAL;
	LRVEL : LREAL;
	LRACC : LREAL;
	LRDEC : LREAL;
	LRJERK : LREAL;
	EDIRECTION : L_TB2P.MC_DIRECTION;
	SCHOMEEXTTP : L_TB2P.MC_TRIGGER_REF;
	XHOMEABSSWITCH : BOOL;
	XSPECIALABORTBEHAVIOR : BOOL;
	LRABORTDEC : LREAL;
	LRABORTJERK : LREAL;
END_VAR
VAR_OUTPUT
	XERROR : BOOL;
	EERRORID : L_TB2P.L_IE1P_Error;
	XFUNBUSY : BOOL;
	XFUNDONE : BOOL;
	XFUNCOMMANDABORTED : BOOL;
	EFUNSTATEACT : L_TB2P.L_MC1P_ABC_State;
	ECONTROLMODE : L_TB2P.L_MC1P_ControlMode;
	XISHOMED : BOOL;
	XHWLIMITSWITCHNEG : BOOL;
	XHWLIMITSWITCHPOS : BOOL;
	XSWLIMITENABLED : BOOL;
	XSWLIMITSWITCHNEG : BOOL;
	XSWLIMITSWITCHPOS : BOOL;
	EAXISTYPE : L_TB2P.L_MC1P_DriveType;
	EAXISSTATE : L_TB2P.L_MC1P_AXIS_STATE;
	XSTOACTIVE : BOOL;
	XREADYFOROPERATION : BOOL;
	XOPERATIONENABLED : BOOL;
	XREADYFORMOTION : BOOL;
	XAXISWARNING : BOOL;
	XAXISERROR : BOOL;
	EAXISERRORID : L_TB2P.L_IE1P_Error;
	XDRIVEWARNING : BOOL;
	XDRIVEERROR : BOOL;
	DWDRIVEERRORID : DWORD;
	LRACTPOS : LREAL;
	LRACTVEL : LREAL;
	LRSETPOSOUT : LREAL;
	LRSETVELOUT : LREAL;
	LRACTFOLLOWINGERROR : LREAL;
	XINPOSITION : BOOL;
	XSTANDSTILLSETVELOCITY : BOOL;
	XSTANDSTILLACTVELOCITY : BOOL;
	XCONSTANTVELOCITY : BOOL;
	XACCELERATING : BOOL;
	XDECELERATING : BOOL;
	XDIRECTIONPOSITIVE : BOOL;
	XDIRECTIONNEGATIVE : BOOL;
	XAXISAVAILABLE : BOOL;
END_VAR
VAR_IN_OUT
	AXIS : AXIS_REF;
END_VAR
END_METHOD

METHOD GET_PAP : POINTER TO L_TB2P_scAP_TM_MotionControl
END_METHOD

METHOD GET_PDATA : POINTER TO L_TS2P_scData_TM_SyncAndCorrectionState
END_METHOD

METHOD GET_PDATASP : POINTER TO L_TS2P_scData_TM_SyncPosBase
END_METHOD

METHOD GET_PPAR : POINTER TO L_TB2P.L_TB2P_scPar_TM_MotionControl
END_METHOD

METHOD GET_PSF : POINTER TO L_TB2P_scSF_TM_MotionControl
END_METHOD

METHOD ADDOFFSET
VAR_INPUT
	ITFTECHMODULE : L_TS2P_ISyncPosBase;
	LRSETPOS : LREAL;
	LRSETVEL : LREAL;
	LRSETOFFSET : LREAL;
	LRSETOFFSETVEL : LREAL;
	ETRAVERSINGRANGE : L_MC1P.L_MC1P_TraversingRange;
	LRCYCLELENGTH : LREAL;
END_VAR
VAR_OUTPUT
	XERROR : BOOL;
	EERRORID : L_IE1P.L_IE1P_Error;
	LRSETPOSOUT : LREAL;
	LRSETVELOUT : LREAL;
END_VAR
END_METHOD

METHOD CLUTCH
VAR_INPUT
	ITFTECHMODULE : L_TS2P_ISyncPosBase;
	XENABLE : BOOL;
	XSYNCIN : BOOL;
	LRSETBASEVELOCITY : LREAL;
	ESYNCMODE : L_TB2P_SyncMode;
	EALLOWEDDIRECTION : L_TB2P_AllowedDirection;
	LRSYNCVEL : LREAL;
	LRSYNCACC : LREAL;
	LRSYNCDEC : LREAL;
	LRSYNCJERK : LREAL;
	LRSYNCINDIST : LREAL;
	LRSYNCOUTDIST : LREAL;
	LRSYNCOUTPOS : LREAL;
	XLOADCLUTCHOFFSET : BOOL;
	LRLOADCLUTCHOFFSET : LREAL;
	LRCYCLICMASTERPOS : LREAL;
	LRCYCLICMASTERVEL : LREAL;
	ETRAVERSINGRANGEMASTER : L_MC1P_TraversingRange;
	LRCYCLELENGTHMASTER : LREAL;
	LRCYCLICAXISPOS : LREAL;
	LRCYCLICAXISVEL : LREAL;
	LRCYCLICAXISACC : LREAL;
	ETRAVERSINGRANGEAXIS : L_MC1P_TraversingRange;
	LRCYCLELENGTHAXIS : LREAL;
END_VAR
VAR_OUTPUT
	XERROR : BOOL;
	EERRORID : L_IE1P.L_IE1P_Error;
	XBUSY : BOOL;
	XDONE : BOOL;
	XSYNCHRONISED : BOOL;
	XACCDECSYNC : BOOL;
	XINBASEVELOCITY : BOOL;
	LRSETPOSOUT : LREAL;
	LRSETVELOUT : LREAL;
	LRSETACCOUT : LREAL;
	LRCLUTCHOFFSETOUT : LREAL;
END_VAR
END_METHOD

METHOD GEARBOX
VAR_INPUT
	ITFTECHMODULE : L_TS2P_ISyncPosBase;
	XENABLE : BOOL;
	LRSETPOSX : LREAL;
	LRSETVELX : LREAL;
	DWNUMERATOR : DWORD;
	DWDENOMINATOR : DWORD;
	LRCYCLELENGTHX : LREAL;
	LRCYCLELENGTHY : LREAL;
	ETRAVERSINGRANGEX : L_MC1P.L_MC1P_TraversingRange;
	ETRAVERSINGRANGEY : L_MC1P.L_MC1P_TraversingRange;
	XLOADGEARBOXPOS : BOOL;
	LRLOADGEARBOXPOS : LREAL;
END_VAR
VAR_OUTPUT
	XERROR : BOOL;
	EERRORID : L_IE1P.L_IE1P_Error;
	LRSETPOSOUT : LREAL;
	LRSETVELOUT : LREAL;
END_VAR
END_METHOD

METHOD OFFSETANDTRIM
VAR_INPUT
	ITFTECHMODULE : L_TS2P_ISyncPosBase;
	XENABLE : BOOL;
	LRSETOFFSET : LREAL;
	XTRIMPOS : BOOL;
	XTRIMNEG : BOOL;
	LRSETTRIMDISTANCE : LREAL;
	ETRIMMODE : L_TS2P_TrimMode;
	XLOADOFFSET : BOOL;
	XRESETTRIMOFFSET : BOOL;
	LRSETVEL : LREAL;
	LRSETACC : LREAL;
	LRSETDEC : LREAL;
	LRSETJERK : LREAL;
	WACTDIRECTION : WORD;
	EALLOWEDDIRECTION : L_TB2P.L_TB2P_AllowedDirection;
	LRCYCMASTERPOS : LREAL;
	LRCYCMASTERVEL : LREAL;
	LRCYCMASTERACC : LREAL;
END_VAR
VAR_OUTPUT
	XERROR : BOOL;
	EERRORID : L_IE1P.L_IE1P_Error;
	XBUSY : BOOL;
	XDONE : BOOL;
	LRSETOFFSETOUTTOTAL : LREAL;
	LRSETOFFSETOUTTOTALVEL : LREAL;
	LRSETOFFSETOUT : LREAL;
	LRSETOFFSETOUTTRIM : LREAL;
END_VAR
END_METHOD

METHOD REQUESTINTERFACE : BOOL
VAR_INPUT
	ID : DINT;
	PITFUNKNOWN : POINTER TO L_UBUP.L_UBUP_IUnknown;
END_VAR
END_METHOD

METHOD CALLFUNCTION
VAR_INPUT
	UIINPUTDATAIDX : UINT;
	UIOUTPUTDATAIDX : UINT;
END_VAR
END_METHOD

METHOD COPYINPUTS : BOOL
VAR_INPUT
	IDX : WORD;
END_VAR
END_METHOD

METHOD COPYOUTPUTS : BOOL
VAR_INPUT
	IDX : WORD;
END_VAR
END_METHOD

METHOD FUNCTIONWASCALLEDTWICE : BOOL
VAR_INPUT
	IDX : WORD;
END_VAR
END_METHOD

METHOD HANDLESTANDARDCALL : BOOL
END_METHOD

METHOD SYNCOUTPUTS
VAR_INPUT
	UICOPYOUTPUTFROMIDX : UINT;
	UICOPYOUTPUTTOIDX : UINT;
END_VAR
END_METHOD

METHOD FB_INIT : BOOL
VAR_INPUT
	BINITRETAINS : BOOL;
	BINCOPYCODE : BOOL;
END_VAR
END_METHOD

METHOD CALL_INTERNALCTRL
END_METHOD

(* ---- L_TS2P_SYNCDRIVEPOS.fb ---- *)
FUNCTION_BLOCK L_TS2P_SYNCDRIVEPOS
VAR_INPUT
	MASTERAXIS : POINTER TO L_MC1P_IAXIS_REF_MASTERVALUES;
	XENABLE : BOOL;
	DWNUMERATOR : DWORD := 1;
	DWDENOMINATOR : DWORD := 1;
	XSYNCIN : BOOL;
	XSYNCOUTINSTANT : BOOL;
	XSYNCINSTANT : BOOL;
	XCLUTCHRELATIVE : BOOL;
	XSYNCPOSRESTORE : BOOL;
	LRSLAVESYNCOUTPOS : LREAL;
	LRSLAVESYNCINDIST : LREAL := 90;
	LRSLAVESYNCOUTDIST : LREAL := 90;
	LRSYNCOUTINSTANTDEC : LREAL := 10000;
	EALLOWEDDIRECTION : L_TB2P_AllowedDirection := L_TB2P_AllowedDirection.both;
	ESYNCMODE : L_TB2P_SyncMode := L_TB2P_SyncMode.ProfGenAbsolute;
	LRSYNCVEL : LREAL := 100;
	LRSYNCACC : LREAL := 1000.0;
	LRSYNCDEC : LREAL := 1000.0;
	LRSYNCJERK : LREAL := 10000000000.0;
	LRSETBASEVELOCITY : LREAL := 0;
	XLOADCLUTCHOFFSET : BOOL := FALSE;
	LRLOADCLUTCHOFFSET : LREAL := 0;
	XTRIMVELOCITYX : BOOL;
	XTRIMVELOCITYY : BOOL;
	LRSETTRIMDISTANCEX : LREAL := 1;
	LRSETTRIMDISTANCEY : LREAL := 1;
	XTRIMPOSX : BOOL;
	XTRIMNEGX : BOOL;
	XTRIMPOSY : BOOL;
	XTRIMNEGY : BOOL;
	XRESETTRIMX : BOOL;
	XRESETTRIMY : BOOL;
	LRSETOFFSETX : LREAL := 0;
	LRSETOFFSETTRIMVELX : LREAL := 10.0;
	LRSETOFFSETTRIMACCX : LREAL := 100.0;
	LRSETOFFSETTRIMDECX : LREAL := 100.0;
	LRSETOFFSETTRIMJERKX : LREAL := 10000.0;
	XLOADOFFSETX : BOOL;
	LRSETOFFSETY : LREAL := 0;
	LRSETOFFSETTRIMVELY : LREAL := 10.0;
	LRSETOFFSETTRIMACCY : LREAL := 100.0;
	LRSETOFFSETTRIMDECY : LREAL := 100.0;
	LRSETOFFSETTRIMJERKY : LREAL := 10000.0;
	XLOADOFFSETY : BOOL;
	XLOADSTARTSLAVEPOS : BOOL := FALSE;
	LRSTARTSLAVEPOS : LREAL;
	XLOADGEARBOXPOS : BOOL;
	LRLOADGEARBOXPOS : LREAL;
	XOPERATIONENABLED : BOOL;
END_VAR
VAR_OUTPUT
	XERROR : BOOL;
	XWARNING : BOOL;
	EERRORID : L_IE1P_Error;
	XBUSY : BOOL;
	LRSETSLAVEPOSOUT : LREAL;
	LRSETSLAVEVELOUT : LREAL;
	LRSETSLAVEACCOUT : LREAL;
	LRSETGEARBOXPOSOUT : LREAL;
	XSYNCOUTDONE : BOOL;
	XSYNCHRONISED : BOOL;
	XACCDECSYNC : BOOL;
	XOFFSETTRIMBUSY : BOOL;
	LROFFSETOUTTOTALVELX : LREAL;
	LROFFSETOUTTOTALVELY : LREAL;
	LROFFSETOUTTRIMX : LREAL;
	LROFFSETOUTTRIMY : LREAL;
	LROFFSETOUTX : LREAL;
	LROFFSETOUTY : LREAL;
	LROFFSETOUTTOTALX : LREAL;
	LROFFSETOUTTOTALY : LREAL;
	LRSETCLUTCHPOS : LREAL;
	LRSETCLUTCHVEL : LREAL;
	LRSETCLUTCHACC : LREAL;
	XBASEVELSYNCHRONISED : BOOL;
	XACCDECBASEVEL : BOOL;
	LROFFSETSYNCPOS : LREAL;
END_VAR
VAR_IN_OUT
	SLAVEAXIS : AXIS_REF;
END_VAR
VAR
	FB_GEARBOXPOSITION : L_MB1P_GearboxPositionInput;
	FB_CLUTCHEXTENDEDBASE : L_TB2P_ClutchExtendedBase;
	FB_AXISCONVERTER : L_MC2P.L_MC2P_AxisConverterBase;
	FB_OFFSETANDTRIMX : L_TS2P_OffsetAndTrim;
	FB_ADDOFFSETCYCLICX : L_MC1P_AddOffsetCyclic;
	FB_OFFSETANDTRIMY : L_TS2P_OffsetAndTrim;
	FB_ADDOFFSETCYCLICY : L_MC1P_AddOffsetCyclic;
	FB_SYNCPOSRESTOREOFFSET : L_TS2P_OffsetAndTrim;
	FB_DIRECTION : L_MC1P_GetDirection;
	LRSETOFFSETMASTER_INT : LREAL;
	LRTRIMDIST_INT : LREAL;
	XTRIMPOS_OLD : BOOL;
	XTRIMNEG_OLD : BOOL;
	XTRIMVEL : BOOL;
	LRTRIMOFFSETDIST : LREAL;
	LRLOADOFFSETMASTER_INT : LREAL := 0;
	LRLOADGEARBOXPOS_INT : LREAL;
	LRSETGEARBOXPOSOUT_INT : LREAL;
	XSETDISABLECLUTCH_INT : BOOL;
	LRLOADTRIMOFFSET_INT : LREAL := 0;
	LRSYNCOUTINSTANTDEC_INT : LREAL := 100000;
	LRSETINTEGRATETRIMVELPOSOUT_INT : LREAL;
	XSYNCPOS_OLD : BOOL;
	XRESETTRIM_OLD : BOOL;
	LRLOADOFFSET_INT : LREAL := 0;
	XSYNCINSTANT_OLD : BOOL;
	XENABLEGEARBOX : BOOL;
	LRSYNCOFFSET : LREAL;
	LRSCALING_INT : LREAL := 1;
	LRGEARBOXSTARTPOSOUT_INT : LREAL;
	DWDENOMINATOR_INT : DWORD := 1;
	XENABLE_OLD : BOOL;
	WAXESMODE : WORD;
	WAXESMODEOLD : WORD;
	LRADDOFFSETPOSOUTY_OLD : LREAL;
	LRADDOFFSETVELOUTY : LREAL;
	LRSETGEARBOXPOSOUTOLD_INT : LREAL;
	LRSETGEARBOXPOSOUTVEL_INT : LREAL;
	LRGETGEARBOXVELIN : LREAL;
	LRGETGEARBOXPOSOUT : LREAL;
	LRGETGEARBOXPOSIN : LREAL;
	LRTASKCYCLE : LREAL;
	XINIT : BOOL := TRUE;
	XCLUTCHDONE_OLD : BOOL;
	XENABLEOLD : BOOL;
	LRSETOFFSETOUTTOTALVELOLD : LREAL;
	SET_AP_LRMASTERVELSTANDSTILLDEADBAND : LREAL;
END_VAR
END_FUNCTION_BLOCK

METHOD CALL_AXESMODE
END_METHOD

METHOD CALL_CALCGEARBOXOUTVELACC
VAR_IN_OUT
	SLAVEAXIS : AXIS_REF;
END_VAR
END_METHOD

METHOD CALL_ERRORHANDLER
END_METHOD

METHOD CALL_FBMETHODS
END_METHOD

METHOD CALL_FBMETHODS_FMDISABLE
END_METHOD

METHOD CALL_FB_ADDOFFSETCYCLICX
END_METHOD

METHOD CALL_FB_ADDOFFSETCYCLICX_INPUT
END_METHOD

METHOD CALL_FB_ADDOFFSETCYCLICY
END_METHOD

METHOD CALL_FB_ADDOFFSETCYCLICY_INPUT
END_METHOD

METHOD CALL_FB_AXISCONVERTER
END_METHOD

METHOD CALL_FB_AXISCONVERTER_INPUT
END_METHOD

METHOD CALL_FB_CLUTCHEXTENDEDBASE
END_METHOD

METHOD CALL_FB_CLUTCHEXTENDEDBASE_INPUT
END_METHOD

METHOD CALL_FB_CLUTCHEXTENDEDBASE_INPUTMASTER
END_METHOD

METHOD CALL_FB_CLUTCHEXTENDEDBASE_INPUTSLAVE
VAR_IN_OUT
	SLAVEAXIS : AXIS_REF;
END_VAR
END_METHOD

METHOD CALL_FB_GEARBOXPOSITION
END_METHOD

METHOD CALL_FB_GEARBOXPOSITION_INPUT
END_METHOD

METHOD CALL_FB_GEARBOXPOSITION_LOADGEARBOXPOS
END_METHOD

METHOD CALL_FB_SYNCPOSRESTOREOFFSET
END_METHOD

METHOD CALL_FB_SYNCPOSRESTOREOFFSET_INPUT
VAR_IN_OUT
	SLAVEAXIS : AXIS_REF;
END_VAR
END_METHOD

METHOD CALL_LOADSLAVESTARTPOS
END_METHOD

METHOD CALL_OFFSETANDTRIMX
END_METHOD

METHOD CALL_OFFSETANDTRIMX_INPUT
END_METHOD

METHOD CALL_OFFSETANDTRIMY
END_METHOD

METHOD CALL_OFFSETANDTRIMY_INPUT
END_METHOD

METHOD CALL_OUTPUT
END_METHOD

METHOD CALL_OUTPUT_CLUTCHSTATE
END_METHOD

METHOD CALL_OUTPUT_OFFSET
END_METHOD

METHOD CALL_RESETCOMMANDS
END_METHOD

METHOD CALL_INIT
VAR_IN_OUT
	SLAVEAXIS : AXIS_REF;
END_VAR
END_METHOD

METHOD GET_DIRECTION
END_METHOD

METHOD GET_GETGEARBOXPOSIN : LREAL
END_METHOD

METHOD GET_GETGEARBOXPOSOUT : LREAL
END_METHOD

METHOD GET_GETGEARBOXVELIN : LREAL
END_METHOD

METHOD GET_GETGEARBOXVELOUT : LREAL
END_METHOD

METHOD GET_LRCLUTCHPOSIN : LREAL
END_METHOD

METHOD GET_LROFFSETADDOFFSETCYCLIC : LREAL
END_METHOD

METHOD SETDISABLECLUTCH : BOOL
VAR_INPUT
	XSETDISABLECLUTCH : BOOL;
END_VAR
END_METHOD

(* ---- L_TS2P_SYNCDRIVEVEL.fb ---- *)
FUNCTION_BLOCK L_TS2P_SYNCDRIVEVEL
VAR_INPUT
	MASTERAXIS : POINTER TO L_MC1P_IAXIS_REF_MASTERVALUES;
	XENABLE : BOOL;
	LRCOUPLINGX : LREAL := 1.0;
	LRCOUPLINGY : LREAL := 1.0;
	XINVERTGEARFACTOR : BOOL;
	XDISABLETOLERANCEINVERTGEARFACTOR : BOOL;
	LRTOLERANCEINVERTGEARFACTOR : LREAL := 0;
	XSYNCIN : BOOL;
	XSYNCOUTINSTANT : BOOL;
	LRSYNCACC : LREAL := 10.0;
	LRSYNCDEC : LREAL := 10.0;
	LRSYNCOUTINSTANTDEC : LREAL := 100.0;
	LRSYNCJERK : LREAL := 1.0;
	XAVOIDVELGAPS : BOOL;
	LRSETOFFSETVEL : LREAL;
	DWMODE : DWORD := 1;
	XTRIMVELOCITYX : BOOL;
	XTRIMVELOCITYY : BOOL;
	LRSETTRIMDISTANCEX : LREAL := 1;
	LRSETTRIMDISTANCEY : LREAL := 1;
	XTRIMPOSX : BOOL;
	XTRIMNEGX : BOOL;
	XTRIMPOSY : BOOL;
	XTRIMNEGY : BOOL;
	XRESETTRIMX : BOOL;
	XRESETTRIMY : BOOL;
	XSYNCVELRESET : BOOL;
	LRSETOFFSETX : LREAL := 0;
	LRSETOFFSETTRIMVELX : LREAL := 10.0;
	LRSETOFFSETTRIMACCX : LREAL := 100.0;
	LRSETOFFSETTRIMDECX : LREAL := 100.0;
	LRSETOFFSETTRIMJERKX : LREAL := 10000.0;
	XLOADOFFSETX : BOOL;
	LRSETOFFSETY : LREAL := 0;
	LRSETOFFSETTRIMVELY : LREAL := 10.0;
	LRSETOFFSETTRIMACCY : LREAL := 100.0;
	LRSETOFFSETTRIMDECY : LREAL := 100.0;
	LRSETOFFSETTRIMJERKY : LREAL := 10000.0;
	XLOADOFFSETY : BOOL;
	EALLOWEDDIRECTION : L_TB2P_AllowedDirection;
	XLOADOFFSET : BOOL;
	XLOADGROUNDVEL : BOOL;
	LRSETGROUNDVEL : LREAL;
	LRGROUNDVELACC : LREAL := 10.0;
	LRGROUNDVELDEC : LREAL := 10.0;
	LRGROUNDVELJERK : LREAL := 1.0;
END_VAR
VAR_OUTPUT
	XERROR : BOOL;
	XWARNING : BOOL;
	EERRORID : L_IE1P_Error;
	XBUSY : BOOL;
	LRSETSLAVEVELOUT : LREAL;
	LRSETSLAVEACCOUT : LREAL;
	XSYNCOUTDONE : BOOL;
	XSYNCHRONISED : BOOL;
	XACCDECSYNC : BOOL;
	XOFFSETTRIMBUSY : BOOL;
	LRPOSOFFSETOUTTRIMX : LREAL;
	LRPOSOFFSETOUTTRIMY : LREAL;
	LRPOSOFFSETOUTX : LREAL;
	LRPOSOFFSETOUTY : LREAL;
	LRPOSOFFSETOUTVELX : LREAL;
	LRVELOFFSET : LREAL;
	LROFFSETOUTTOTALX : LREAL;
	LROFFSETOUTTOTALY : LREAL;
	LROFFSETOUTTOTALVELX : LREAL;
	LROFFSETOUTTOTALVELY : LREAL;
	XBASEVELSYNCHRONISED : BOOL;
	XACCDECBASEVEL : BOOL;
	XBASEVELSYNCOUTDONE : BOOL;
	XINVERTGEARFACTORACTIVE : BOOL;
END_VAR
VAR_IN_OUT
	SLAVEAXIS : AXIS_REF;
END_VAR
VAR
	XENABLE_OLD : BOOL;
	ESTATE : L_TF1P_States := L_TF1P_States.INIT;
	ESTATE_OLD : L_TF1P_States := L_TF1P_States.INIT;
	XSTATEENTRY : BOOL;
	FB_CONVAXISV : L_MC2P_ConvAxisV;
	FB_INVERTGEARFACTOR : L_TS2P_InvertGearfactor;
	XACCDECSYNC_OLD : BOOL;
	XSYNCVEL_OLD : BOOL;
	XOPEN_OLD : BOOL;
	LRSETVELTRIM : LREAL;
	XSETDISABLECLUTCH_INT : BOOL;
	SETPOSITIONFORSYNCOLD : LREAL := 0;
	XINITFB_CLUTCHV : BOOL;
	FB_CLUTCHV : L_MC2P_ClutchVelocity;
	XINVERTGEARFACTORACTIVE_OLD : BOOL;
	LRSETGROUNDVEL_INT : LREAL;
	FB_OFFSETANDTRIMX : L_TS2P_OffsetAndTrim;
	FB_VELOCITYOFFSET : L_MC1P_RampGenerator;
	FB_OFFSETANDTRIMY : L_TS2P_OffsetAndTrim;
	FB_RAMPGENGROUNDVEL : L_MC1P_RampGenerator;
	FB_DIRECTION : L_MC1P_GetDirection;
END_VAR
END_FUNCTION_BLOCK

METHOD CALL_ERRORHANDLER
END_METHOD

METHOD CALL_FBMETHODS
END_METHOD

METHOD CALL_FBMETHODS_FMDISABLE
END_METHOD

METHOD CALL_FB_CLUTCHV
END_METHOD

METHOD CALL_FB_CLUTCHV_INPUT
END_METHOD

METHOD CALL_FB_CLUTCHV_PAR
END_METHOD

METHOD CALL_FB_CONVAXISV
END_METHOD

METHOD CALL_FB_CONVAXISV_INPUT
END_METHOD

METHOD CALL_FB_INVERTGEARFACTOR
END_METHOD

METHOD CALL_FB_INVERTGEARFACTOR_INPUT
END_METHOD

METHOD CALL_FB_RAMPGENGROUNDVEL
END_METHOD

METHOD CALL_FB_RAMPGENGROUNDVEL_INPUT
END_METHOD

METHOD CALL_FB_VELOCITYOFFSET
END_METHOD

METHOD CALL_FB_VELOCITYOFFSET_INPUT
END_METHOD

METHOD CALL_OFFSETANDTRIMX
END_METHOD

METHOD CALL_OFFSETANDTRIMX_INPUT
END_METHOD

METHOD CALL_OFFSETANDTRIMY
END_METHOD

METHOD CALL_OFFSETANDTRIMY_INPUT
END_METHOD

METHOD CALL_OUTPUT
END_METHOD

METHOD CALL_OUTPUT_SETSLAVEOUT
END_METHOD

METHOD CALL_RESETCOMMANDS
END_METHOD

METHOD CALL_RESETFM
END_METHOD

METHOD CALL_RESETOUTPUT
END_METHOD

METHOD CALL_STATEMASHINE
END_METHOD

METHOD GET_DIRECTION
END_METHOD

METHOD GET_CLUTCHVELOUT : LREAL
END_METHOD

METHOD GET_GETGEARBOXVELIN : LREAL
END_METHOD

METHOD GET_GETGEARBOXVELOUT : LREAL
END_METHOD

METHOD SETDISABLECLUTCH : BOOL
VAR_INPUT
	XSETDISABLECLUTCH : BOOL;
END_VAR
END_METHOD

METHOD CALL_S000_CYCLIC
END_METHOD

METHOD CALL_S001_INIT
END_METHOD

METHOD CALL_S010_READY
END_METHOD

METHOD CALL_S998_ERROR
END_METHOD

(* ---- L_TS2P_SYNCPOSBASE.fb ---- *)
FUNCTION_BLOCK L_TS2P_SYNCPOSBASE EXTENDS L_TB2P_TechModuleBase
VAR_INPUT
	XUSEORIGINAL : BOOL;
	XENABLE : BOOL;
	XENABLEOPERATION : BOOL;
	XRESETERROR : BOOL;
	XQSPAPPLICATION : BOOL;
	XABORT : BOOL;
	XJOGPOS : BOOL;
	XJOGNEG : BOOL;
	XHOMEEXECUTE : BOOL;
	LROVERRIDE : LREAL := 1;
	SCCTRLBASICMOTION : L_TB2P_scCtrlBasicMotion;
	SCPAR : L_TS2P_scPar_SyncPosBase;
	SCACCESSPOINTS : L_TS2P_scAP_SyncPosBase;
	MASTERVALUES : L_MC1P_IAXIS_REF_MASTERVALUES;
	XSYNCIN : BOOL;
	XSYNCPOSRESTORE : BOOL;
	LRSETBASEVEL : LREAL;
	LRSETOFFSETPOS : LREAL;
	XTRIMPOS : BOOL;
	XTRIMNEG : BOOL;
	XTRIMRESET : BOOL;
END_VAR
VAR_OUTPUT
	XREADYFOROPERATION : BOOL;
	XOPERATIONENABLED : BOOL;
	XREADYFORMOTION : BOOL;
	XERROR : BOOL;
	XWARNING : BOOL;
	EERRORID : L_IE1P_Error;
	XSTOACTIVE : BOOL;
	XQSPACTIVE : BOOL;
	XABORTBUSY : BOOL;
	XABORTDONE : BOOL;
	XJOGGINGBUSY : BOOL;
	XHOMINGBUSY : BOOL;
	XHOMINGDONE : BOOL;
	XISHOMED : BOOL;
	ETMSTATE : L_TB2P_States;
	SCSTATUSBASICMOTION : L_TB2P_scStatusBasicMotion;
	LRACTVEL : LREAL;
	LRSETVELOUT : LREAL;
	LRACTPOS : LREAL;
	LRSETPOSOUT : LREAL;
	LRACTFOLLOWINGERROR : LREAL;
	SCSIGNALFLOW : L_TS2P_scSF_SyncPosBase;
	XSYNCHRONISED : BOOL;
	XACCDECSYNC : BOOL;
	XOFFSETTRIMACTIVE : BOOL;
	XBASEVELOCITYACTIVE : BOOL;
	LROFFSETTOTAL : LREAL;
END_VAR
VAR_IN_OUT
	AXIS : AXIS_REF;
END_VAR
VAR
	XINTERNALCONTROLACTIVE_OLD : BOOL;
	ITFCONNECTORSYNCPOS : L_TS2P_IConnectorSyncPos;
	_XCONNECTORVALID : BOOL;
	TM_INT : L_TS2P_TM_SyncPosBase;
	SCPAR_INT : L_TS2P_scPar_SyncPosBase;
	SCDATA_INT : L_TS2P_scData_TM_SyncPosBase;
	XUSEORIGINAL_OLD : BOOL;
	_UICALLMFUNIDXINPUT : UINT := 1;
	_UICALLMFUNIDXOUTPUT : UINT := 1;
	_MCCALL : L_UM1P_MCCall := STRUCT(itfMCCall := THIS^);
	_ASCINPUT : ARRAY [1.._MCCall.c_BufferDepthInput] OF L_TS2P_SyncPosBaseIn;
	_ASCOUTPUT : ARRAY [1.._MCCall.c_BufferDepthOutput] OF L_TS2P_SyncPosBaseOut;
	_ASCPARCORE : ARRAY [1.._MCCall.c_BufferDepthInput] OF L_TS2P_scPar_SyncPosBase;
	_ASCACCESSPOINTSCORE : ARRAY [1.._MCCall.c_BufferDepthInput] OF L_TS2P_scAP_SyncPosBase;
	_ASCSIGNALFLOWCORE : ARRAY [1.._MCCall.c_BufferDepthOutput] OF L_TS2P_scSF_SyncPosBase;
	_SCINPUTVISU : L_TS2P_SyncPosBaseIn;
	_PSCINPUTVISU : POINTER TO L_TS2P_SyncPosBaseIn := ADR(_scInputVisu);
	_PSCOUTPUTVISU : POINTER TO L_TS2P_SyncPosBaseOut := ADR(_ascOutput[1]);
	_PSCDATAVISU : POINTER TO L_TS2P_scData_TM_SyncPosBase := ADR(scData_int);
	_PSCPARVISU : POINTER TO L_TS2P_scPar_SyncPosBase := ADR(scPar_int);
	_PSCAPVISU : POINTER TO L_TS2P_scAP_SyncPosBase;
	_PSCSFVISU : POINTER TO L_TS2P_scSF_SyncPosBase;
	ITFBASICMOTIONBASE : L_TB2P.L_TB2P_IBasicMotionBase;
	ITFITECHMODULEINTERNAL : L_TB2P_ITechModuleInternal;
	ITFSYNCPOSEXTENSION : L_TS2P_ISyncPosBase;
	LRJERKDEC : LREAL;
	LRJOGGINGJERKDEC : LREAL;
	REMAININGTIMEOFPROFILE : LREAL;
	REMAININGTIMEOFPROFILEAVAILABLE : BOOL;
END_VAR
END_FUNCTION_BLOCK

METHOD CALL_ABC
VAR_INPUT
	ITFTECHMODULE : L_TB2P.L_TB2P_IBasicMotionBase;
	XQSPAPPLICATION : BOOL;
	XHALT : BOOL;
	XABORT : BOOL;
	XHOMEEXECUTE : BOOL;
	XJOGPOS : BOOL;
	XJOGNEG : BOOL;
	XFINISHPOSITIONING : BOOL;
	XMOVEVELEXECUTE : BOOL;
	XMOVEABSEXECUTE : BOOL;
	XMOVERELEXECUTE : BOOL;
	XENABLEOPERATION : BOOL;
	XRESETERROR : BOOL;
	XENABLEPOSITIVE : BOOL;
	XENABLENEGATIVE : BOOL;
	XDISABLESWLIMIT : BOOL;
	LROVERRIDE : LREAL;
	LROVERRIDEACC : LREAL;
	LROVERRIDEJERK : LREAL;
	XRESETHOMEPOSITION : BOOL;
	XCONTINUOUSUPDATE : BOOL;
	LRPOS_DIST : LREAL;
	LRVEL : LREAL;
	LRACC : LREAL;
	LRDEC : LREAL;
	LRJERK : LREAL;
	EDIRECTION : L_TB2P.MC_DIRECTION;
	SCHOMEEXTTP : L_TB2P.MC_TRIGGER_REF;
	XHOMEABSSWITCH : BOOL;
	XSPECIALABORTBEHAVIOR : BOOL;
	LRABORTDEC : LREAL;
	LRABORTJERK : LREAL;
END_VAR
VAR_OUTPUT
	XERROR : BOOL;
	EERRORID : L_TB2P.L_IE1P_Error;
	XFUNBUSY : BOOL;
	XFUNDONE : BOOL;
	XFUNCOMMANDABORTED : BOOL;
	EFUNSTATEACT : L_TB2P.L_MC1P_ABC_State;
	ECONTROLMODE : L_TB2P.L_MC1P_ControlMode;
	XISHOMED : BOOL;
	XHWLIMITSWITCHNEG : BOOL;
	XHWLIMITSWITCHPOS : BOOL;
	XSWLIMITENABLED : BOOL;
	XSWLIMITSWITCHNEG : BOOL;
	XSWLIMITSWITCHPOS : BOOL;
	EAXISTYPE : L_TB2P.L_MC1P_DriveType;
	EAXISSTATE : L_TB2P.L_MC1P_AXIS_STATE;
	XSTOACTIVE : BOOL;
	XREADYFOROPERATION : BOOL;
	XOPERATIONENABLED : BOOL;
	XREADYFORMOTION : BOOL;
	XAXISWARNING : BOOL;
	XAXISERROR : BOOL;
	EAXISERRORID : L_TB2P.L_IE1P_Error;
	XDRIVEWARNING : BOOL;
	XDRIVEERROR : BOOL;
	DWDRIVEERRORID : DWORD;
	LRACTPOS : LREAL;
	LRACTVEL : LREAL;
	LRSETPOSOUT : LREAL;
	LRSETVELOUT : LREAL;
	LRACTFOLLOWINGERROR : LREAL;
	XINPOSITION : BOOL;
	XSTANDSTILLSETVELOCITY : BOOL;
	XSTANDSTILLACTVELOCITY : BOOL;
	XCONSTANTVELOCITY : BOOL;
	XACCELERATING : BOOL;
	XDECELERATING : BOOL;
	XDIRECTIONPOSITIVE : BOOL;
	XDIRECTIONNEGATIVE : BOOL;
	XAXISAVAILABLE : BOOL;
END_VAR
VAR_IN_OUT
	AXIS : AXIS_REF;
END_VAR
END_METHOD

METHOD GET_PAP : POINTER TO L_TB2P_scAP_TM_MotionControl
END_METHOD

METHOD GET_PDATA : POINTER TO L_TS2P_scData_TM_SyncPosBase
END_METHOD

METHOD GET_PPAR : POINTER TO L_TB2P.L_TB2P_scPar_TM_MotionControl
END_METHOD

METHOD GET_PSF : POINTER TO L_TB2P_scSF_TM_MotionControl
END_METHOD

METHOD ADDOFFSET
VAR_INPUT
	ITFTECHMODULE : L_TS2P_ISyncPosBase;
	LRSETPOS : LREAL;
	LRSETVEL : LREAL;
	LRSETOFFSET : LREAL;
	LRSETOFFSETVEL : LREAL;
	ETRAVERSINGRANGE : L_MC1P.L_MC1P_TraversingRange;
	LRCYCLELENGTH : LREAL;
END_VAR
VAR_OUTPUT
	XERROR : BOOL;
	EERRORID : L_IE1P.L_IE1P_Error;
	LRSETPOSOUT : LREAL;
	LRSETVELOUT : LREAL;
END_VAR
END_METHOD

METHOD CLUTCH
VAR_INPUT
	ITFTECHMODULE : L_TS2P_ISyncPosBase;
	XENABLE : BOOL;
	XSYNCIN : BOOL;
	LRSETBASEVELOCITY : LREAL;
	ESYNCMODE : L_TB2P_SyncMode;
	EALLOWEDDIRECTION : L_TB2P_AllowedDirection;
	LRSYNCVEL : LREAL;
	LRSYNCACC : LREAL;
	LRSYNCDEC : LREAL;
	LRSYNCJERK : LREAL;
	LRSYNCINDIST : LREAL;
	LRSYNCOUTDIST : LREAL;
	LRSYNCOUTPOS : LREAL;
	XLOADCLUTCHOFFSET : BOOL;
	LRLOADCLUTCHOFFSET : LREAL;
	LRCYCLICMASTERPOS : LREAL;
	LRCYCLICMASTERVEL : LREAL;
	ETRAVERSINGRANGEMASTER : L_MC1P_TraversingRange;
	LRCYCLELENGTHMASTER : LREAL;
	LRCYCLICAXISPOS : LREAL;
	LRCYCLICAXISVEL : LREAL;
	LRCYCLICAXISACC : LREAL;
	ETRAVERSINGRANGEAXIS : L_MC1P_TraversingRange;
	LRCYCLELENGTHAXIS : LREAL;
END_VAR
VAR_OUTPUT
	XERROR : BOOL;
	EERRORID : L_IE1P.L_IE1P_Error;
	XBUSY : BOOL;
	XDONE : BOOL;
	XSYNCHRONISED : BOOL;
	XACCDECSYNC : BOOL;
	XINBASEVELOCITY : BOOL;
	LRSETPOSOUT : LREAL;
	LRSETVELOUT : LREAL;
	LRSETACCOUT : LREAL;
	LRCLUTCHOFFSETOUT : LREAL;
END_VAR
END_METHOD

METHOD GEARBOX
VAR_INPUT
	ITFTECHMODULE : L_TS2P_ISyncPosBase;
	XENABLE : BOOL;
	LRSETPOSX : LREAL;
	LRSETVELX : LREAL;
	DWNUMERATOR : DWORD;
	DWDENOMINATOR : DWORD;
	LRCYCLELENGTHX : LREAL;
	LRCYCLELENGTHY : LREAL;
	ETRAVERSINGRANGEX : L_MC1P.L_MC1P_TraversingRange;
	ETRAVERSINGRANGEY : L_MC1P.L_MC1P_TraversingRange;
	XLOADGEARBOXPOS : BOOL;
	LRLOADGEARBOXPOS : LREAL;
END_VAR
VAR_OUTPUT
	XERROR : BOOL;
	EERRORID : L_IE1P.L_IE1P_Error;
	LRSETPOSOUT : LREAL;
	LRSETVELOUT : LREAL;
END_VAR
END_METHOD

METHOD OFFSETANDTRIM
VAR_INPUT
	ITFTECHMODULE : L_TS2P_ISyncPosBase;
	XENABLE : BOOL;
	LRSETOFFSET : LREAL;
	XTRIMPOS : BOOL;
	XTRIMNEG : BOOL;
	LRSETTRIMDISTANCE : LREAL;
	ETRIMMODE : L_TS2P_TrimMode;
	XLOADOFFSET : BOOL;
	XRESETTRIMOFFSET : BOOL;
	LRSETVEL : LREAL;
	LRSETACC : LREAL;
	LRSETDEC : LREAL;
	LRSETJERK : LREAL;
	WACTDIRECTION : WORD;
	EALLOWEDDIRECTION : L_TB2P.L_TB2P_AllowedDirection;
	LRCYCMASTERPOS : LREAL;
	LRCYCMASTERVEL : LREAL;
	LRCYCMASTERACC : LREAL;
END_VAR
VAR_OUTPUT
	XERROR : BOOL;
	EERRORID : L_IE1P.L_IE1P_Error;
	XBUSY : BOOL;
	XDONE : BOOL;
	LRSETOFFSETOUTTOTAL : LREAL;
	LRSETOFFSETOUTTOTALVEL : LREAL;
	LRSETOFFSETOUT : LREAL;
	LRSETOFFSETOUTTRIM : LREAL;
END_VAR
END_METHOD

METHOD REQUESTINTERFACE : BOOL
VAR_INPUT
	ID : DINT;
	PITFUNKNOWN : POINTER TO L_UBUP.L_UBUP_IUnknown;
END_VAR
END_METHOD

METHOD CALLFUNCTION
VAR_INPUT
	UIINPUTDATAIDX : UINT;
	UIOUTPUTDATAIDX : UINT;
END_VAR
END_METHOD

METHOD COPYINPUTS : BOOL
VAR_INPUT
	IDX : WORD;
END_VAR
END_METHOD

METHOD COPYOUTPUTS : BOOL
VAR_INPUT
	IDX : WORD;
END_VAR
END_METHOD

METHOD FUNCTIONWASCALLEDTWICE : BOOL
VAR_INPUT
	IDX : WORD;
END_VAR
END_METHOD

METHOD HANDLESTANDARDCALL : BOOL
END_METHOD

METHOD SYNCOUTPUTS
VAR_INPUT
	UICOPYOUTPUTFROMIDX : UINT;
	UICOPYOUTPUTTOIDX : UINT;
END_VAR
END_METHOD

METHOD FB_INIT : BOOL
VAR_INPUT
	BINITRETAINS : BOOL;
	BINCOPYCODE : BOOL;
END_VAR
END_METHOD

METHOD CALL_INTERNALCTRL
END_METHOD

(* ---- L_TS2P_SYNCRONISEDOVERRIDE.fb ---- *)
FUNCTION_BLOCK L_TS2P_SYNCRONISEDOVERRIDE
VAR_INPUT
	XENABLE : BOOL;
	XSYNCHRONISED : BOOL;
	XEXECUTEGAP : BOOL;
	XAUXEXECUTEGAP : BOOL;
	LRSYNCOVERRIDE : LREAL := 1;
	LRCYCMASTERPOS : LREAL;
	LRCYCMASTERVEL : LREAL;
	LRCYCMASTERACC : LREAL;
	LRCYCSLAVEPOS : LREAL;
	LRCYCSLAVEVEL : LREAL;
	LRCYCSLAVEACC : LREAL;
	LRACC : LREAL;
	LRDEC : LREAL;
	LRJERK : LREAL;
	LRTASKCYLCETIME : LREAL := 0.001;
END_VAR
VAR_OUTPUT
	XBUSY : BOOL;
	XERROR : BOOL;
	EERRORID : L_IE1P_Error;
	XOVERRIDELIMITED : BOOL;
	XEXECUTEGAPOUT : BOOL;
	XAUXEXECUTEGAPOUT : BOOL;
	LRSETPOS : LREAL;
	LRSETVEL : LREAL;
	LRSETACC : LREAL;
	XSYNCOVERRIDEACTIVE : BOOL;
	XRAMPGENBUSY : BOOL;
END_VAR
VAR
	XENABLE_OLD : BOOL;
	XEXECUTEGAP_OLD : BOOL;
	XAUXEXECUTEGAP_OLD : BOOL;
	LRSYNCOVERRIDE_INT : LREAL := 1;
	LRSYNCOVERRIDE_LOCK : LREAL;
	LRADDOVERRIDE_LOCK : LREAL;
	WSTATE : WORD := 0;
	LROFFSETPOS_INT : LREAL;
	LROFFSETVEL_INT : LREAL;
	LROFFSETACC_INT : LREAL;
	LROFFSETVEL_OLD : LREAL;
	LRVELTARGET : LREAL;
	LRVELSTART : LREAL;
	FB_RAMPGENERATOR1 : L_MC1P_RampGenerator;
	C_LRCYCLELENGTHMASTER : LREAL := (16#4FFFFFFFFFFFFFFF * 1E-08);
END_VAR
END_FUNCTION_BLOCK

METHOD CALL_ERRORHANDLER
END_METHOD

METHOD CALL_FB_RAMPGENERATOR1
END_METHOD

METHOD CALL_OUTPUTS
END_METHOD

METHOD CALL_RESETCOMMANDS
END_METHOD

METHOD CALL_RESETOUTPUTS
END_METHOD

METHOD CALL_STATEMACHINE
END_METHOD

(* ---- L_TS2P_TM_CROSSCUTTERBASE.fb ---- *)
FUNCTION_BLOCK L_TS2P_TM_CROSSCUTTERBASE EXTENDS L_TB2P_SyncMotionControl
VAR_OUTPUT
	PAP : POINTER TO L_TS2P_scAP_TM_CrossCutterHigh;
	PSF : POINTER TO L_TS2P_scSF_TM_CrossCutterHigh;
	PPAR : POINTER TO L_TS2P_scPar_TM_CrossCutterHigh := ADR(scPar_int);
	PPARBASE : POINTER TO L_TS2P_scPar_TM_CrossCutterBaseExtension := ADR(scPar_int);
END_VAR
VAR
	TM_CROSSCUTTERBASECONFIG : L_TB2P_ModuleHandlerConfig;
	PSCINPUT : POINTER TO L_TS2P_CrossCutterStateIn;
	PSCOUTPUT : POINTER TO L_TS2P_CrossCutterStateOut;
	LROFFSET : LREAL;
	LROFFSETTRIM : LREAL;
	XSYNCOUTINSTANT_INT : BOOL;
	PMASTERAXIS : POINTER TO _AXIS_REF_REAL;
	LRCUTTINGANGLE_INT : LREAL;
	SCPAR_INT : L_TS2P_scPar_TM_CrossCutterHigh;
	LRSLAVEMAXVEL_INT : LREAL;
	LRSLAVEMAXACC_INT : LREAL;
	XCUTTINGBUSY_INT : BOOL;
	XACCDECSYNC_INT : BOOL;
	XCCMOVEABSEXECUTE_INT : BOOL;
	LRCCPOS_DIST_INT : LREAL;
	BYSETTOOLNOOUT : BYTE;
	BYSETAREAOUT : BYTE;
	LRSETXPOSOUT : LREAL;
	LRSETXVELOUT : LREAL;
	LRSETXACCOUT : LREAL;
	LRSLAVEMAXVEL : LREAL;
	LRSLAVEMAXACC : LREAL;
	LRMASTERVEL : LREAL;
	LRMASTERVEL_OLD : LREAL;
	LRMASTERVEL_OLD2 : LREAL;
	LRMASTERPOS_OLD : LREAL;
	LRACTMASTERPOS_OLD : LREAL;
	XMASTERAXISENABLED : BOOL;
	XMASTERAXISENABLED_OLD : BOOL;
	XCUTTINGACTIVE_OLD : BOOL;
	XRESETTRIMOFFSET_OLD : BOOL;
	XENABLECONTROLSETVALUES_OLD : BOOL;
	XINPARKPOS_OLD : BOOL;
	XMASTERISSTANDSTILL : BOOL;
	XNEXTTOOLDIRECTIONPOSITIV : BOOL := TRUE;
	ECUTTINGPROCESSSTATE : L_TB2P_States := L_TB2P_States.DISABLED;
	_XCALLCALLUTTINGPROCESSAGAIN : BOOL;
	BYPOSITIONINGSTATE : BYTE := 0;
	BYMASTEROFFSETSTEPPER : BYTE := 0;
	BYTOOLCIRCARRAYPREPARED : BYTE;
	XMASTERIS_FREEENCODER : BOOL;
	XEXECUTETRANSITIONCYCLES : BOOL;
	XINVALIDCROSSCUTTERPARAMETRS : BOOL;
	XINVALIDCUTTINGPARAMETRS : BOOL;
	XMASTERNOTROTATIVE : BOOL;
	XWARNINGINVALIDPRODUCTLENGTH : BOOL;
	XINVALIDPRODUCTLENGTH : BOOL;
	XINVALIDCUTTINGANGLE : BOOL;
	XSLAVEOUTOFSCALE : BOOL;
	XERRORSLAVENOTINPARKPOS : BOOL;
	XMASTEROUTOFSCALE : BOOL;
	XSLAVERECEIVEDGAPS : BOOL;
	XINVALIDCAMSELECTED : BOOL;
	XWARNINGINVALIDCAMSELECTED : BOOL;
	XWARNINGDIRECTIONDISABLEDSYNCINT : BOOL;
	XWARNINGAXISNOTHOMED4SYNCIN : BOOL;
	ILOOPCNTR : INT;
	UIVARTEMP : UINT;
	IVARTEMP : INT;
	LRVARTEMP : LREAL;
	LRVARTEMP2 : LREAL;
	LRVARTEMP3 : LREAL;
	LRVARTEMP4 : LREAL;
	LRTEMPSTOPLENGTH : LREAL;
	LRTEMPSTARTLENGTH : LREAL;
	LRXDISTINPARKPOS : LREAL;
	XXPOSSYNCRONISEDMASTERPOS : BOOL;
	XCUTTINGPARISCHANGED : BOOL;
	XCAMDIRECTCHANGE_LOCK : BOOL;
	LRSETMASTERTRIMOFFSET_INT : LREAL;
	LRSETOFFSETMASTER_LOCK : LREAL;
	LRSETMASTERTRIMOFFSET_LOCK : LREAL;
	LRSETMASTERTRIMOFFSET_SAVE : LREAL;
	_LROFFSETTOTAL_OLD : LREAL;
	WLENGTHCALCULATORMODE : WORD := 2;
	LRACTMASTERPOSSTART : LREAL;
	LRLENGTHCALCULATOR : LREAL;
	LROVERSPEEDUPPERLIMIT : LREAL := 2;
	ECUTTINGMODE_LOCK : L_TS2P_CuttingModeState;
	BYCAMCONTINUOUSNO_LOCK : BYTE := 1;
	BYNUMOFTOOLS_LOCK : BYTE;
	LRPRODUCTLENGTH_LOCK : LREAL;
	LRPRODUCTLENGTH_LOCK_OLD : LREAL;
	LRCUTLENGTH_LOCK : LREAL;
	LROSCILLATION_LOCK : LREAL := 0;
	LROVERSPEED_LOCK : LREAL;
	LROVERSPEEDFACTOR_LOCK : LREAL;
	LROVERSPEEDFACTOR_LOCK_OLD : LREAL;
	LRCUTTINGANGLE_LOCK : LREAL;
	LRSCALINGMASTER_LOCK : LREAL := 1;
	LRTOOLTOOLDIST_LOCK : LREAL;
	LRTOOLTOOLCIRCUMFERENCEDIST_LOCK : LREAL;
	LRCIRCUMFERENCE_LOCK : LREAL;
	LRCIRCUMFERENCEINV_LOCK : LREAL;
	XHOLDINPARKPOS_LOCK : BOOL;
	LRFACTOR_ANGLETOSLAVEUNITS_LOCK : LREAL;
	LRFACTOR_ANGLETOMASTERUNITS_LOCK : LREAL;
	LRFACTOR_SLAVEUNITSTOMASTERUNITS_LOCK : LREAL;
	LRFACTOR_MASTERUNITSTOSLAVEUNITS_LOCK : LREAL;
	LRFACTOR_PRODUCTUNITSTOMASTERUNITS_LOCK : LREAL;
	LRFACTOR_PRODUCTUNITSTOMASTERUNITSINV_LOCK : LREAL;
	LRFACTOR_PRODUCTUNITSTOMASTERUNITSINV_OLD : LREAL;
	XFIRSTCUT : BOOL;
	XCONTINUOUSMODE : BOOL := TRUE;
	BYSETCAMTABLENO : BYTE;
	BYREQUESTSSETCAMTABLE : BYTE;
	BYREQUESTSSETCAMTABLE_OLD : BYTE;
	SCSYNCSTARTLENGTH : L_MC2P_CamDataXYVA;
	SCSYNCSTOPLENGTH : L_MC2P_CamDataXYVA;
	SCASYNCLENGTH : L_MC2P_CamDataXYVA;
	SCSTARTLENGTH : L_MC2P_CamDataXYVA;
	SCSTOPLENGTH : L_MC2P_CamDataXYVA;
	LRSTANDSTILLLENGTH : LREAL;
	LRY_START : LREAL := 0;
	LRY_PARK : LREAL := 180;
	LRY_END : LREAL := 360;
	LRX_START : LREAL := 0;
	LRX_ENDSYNCPOS : LREAL := 10;
	LRX_STARTPARKPOS : LREAL := 180;
	LRX_ENDPARKPOS : LREAL := 180;
	LRX_STARTSYNCPOS : LREAL := 350;
	LRX_END : LREAL := 360;
	LRY_END_PREVIOUSLY : LREAL := 360;
	LRY_CUTLENGTHCALCULATOR : LREAL := 360;
	LROVERSPEED_LOCK_PREVIOUSLY : LREAL;
	FM_CAMCREATOR_START : L_TS2P_CamCreator;
	FM_CAMCREATOR_STOP : L_TS2P_CamCreator;
	FM_CAMCREATOR_CONTINUOUS : ARRAY [1..2] OF L_TS2P_CamCreator;
	FM_CAMCREATOR_STANDSTILL : L_TS2P_CamCreator;
	CAM_START_P : ARRAY [0..3] OF L_MC2P_CamDataXYVA;
	CAM_STOP_P : ARRAY [0..3] OF L_MC2P_CamDataXYVA;
	CAM_CONTINUOUS_P : ARRAY [1..2] OF ARRAY [0..3] OF L_MC2P_CamDataXYVA;
	CAM_STOPSTART_P : ARRAY [1..2] OF ARRAY [0..5] OF L_MC2P_CamDataXYVA;
	CAM_STANDSTILL_P : ARRAY [0..1] OF L_MC2P_CamDataXYVA;
	CAMTABLEATFLEXCAM : MC_CAM_REF;
	LRYOFFSET : LREAL;
	LRENDOFPROFILEWINDOWSIZE : LREAL := 0;
	_FC_XMASTERABSOLUTE : BOOL;
	_FC_XSLAVEABSOLUTE : BOOL;
	_FC_XPERIODIC : BOOL;
	_FC_XTRIMMASTERNEG : BOOL;
	_FC_XTRIMMASTERPOS : BOOL;
	_FC_LRSETOFFSETMASTER : LREAL;
	_FC_LRSETOFFSETSLAVE : LREAL;
	_FC_EPOSCTRLDIRECTION : L_MC2P.L_MC2P_ReverseCtrlDirection;
	_FC_EOFFSETMODEMASTER : L_MC2P.L_MC2P_OffsetMode;
	_FC_EOFFSETMODESLAVE : L_MC2P.L_MC2P_OffsetMode;
	_FC_XHOLDPROFGENMASTER : BOOL;
	_FC_ESYNCMODE : L_MC2P.L_MC2P_ClutchMode;
	_FC_ESYNCDIRECTION : L_MC2P.L_MC2P_ClutchDirection;
	_FC_LRMASTERSYNCINDIST : LREAL;
	_FC_LRMASTERSYNCINPOS : LREAL;
	_FC_LRMASTERSYNCOUTDIST : LREAL;
	_FC_LRSLAVESYNCOUTPOS : LREAL;
	_FC_LRSYNCINTIME : LREAL;
	_FC_LRSYNCOUTTIME : LREAL;
	_FC_LRSYNCOUTINSTANTDEC : LREAL;
	_FC_XENABLE : BOOL;
	_FC_XSYNCPOS : BOOL;
	_FC_XSYNCCAM : BOOL;
	_FC_XDIRECTCHANGE : BOOL;
	_FC_XSYNCOUTINSTANT : BOOL;
	_XCUTTINGACTIVECUTDONE : BOOL;
	_FC_LRSYNCCAMVEL : LREAL;
	_FC_LRSYNCCAMACC : LREAL;
	_FC_LRSYNCCAMDEC : LREAL;
	_FC_LRSYNCCAMJERK : LREAL;
	_FC_LRSETXPOSOUT : LREAL;
	_FC_LRSETXVELOUT : LREAL;
	_FC_LRSETXACCOUT : LREAL;
	_FC_LRSETYPOSOUT : LREAL;
	_FC_LRSETYVELOUT : LREAL;
	_FC_LRSETYACCOUT : LREAL;
	_FC_LRSETSLAVEPOSOUT : LREAL;
	_FC_LRSETSLAVEVELOUT : LREAL;
	_FC_LRSETSLAVEACCOUT : LREAL;
	_FC_XENDOFPROFILE : BOOL;
	_FC_XACCDECSYNC : BOOL;
	_FC_XSYNCHRONISED : BOOL;
	_FC_LRSETOFFSETMASTEROUT : LREAL;
	_FC_XENDOFCYCLE : BOOL;
	_FC_LRSETXPOS : LREAL;
	_FC_XCAMSYNCHRONISED : BOOL;
	_FC_XDONE : BOOL;
	_FC_XBUSY : BOOL;
	_FC_LRSETMASTERTRIMOFFSETOUT : LREAL;
	_FC_XENDOFPROFNEGATIVE : BOOL;
	_FC_LWENDOFPROFILECHECKSUM : LWORD;
	FM_FLEXCAMHIGH : L_MC2P_FlexCamHigh;
	FB_CONTROLSETVALUES : L_MC1P_ControlSetValues := STRUCT(eSetValueMode := L_MC1P_SetValueMode.Pos);
	L_MB1P_DIFFERENTIATE1 : L_MC2P_Differentiate;
	XINTERNALERROR : BOOL;
	WINTERNALERRORID : WORD;
	LWTCHECKSUM_INT : LWORD;
END_VAR
END_FUNCTION_BLOCK

METHOD CALL_ALLOCPOINTADR
END_METHOD

METHOD CALL_CTRLREQACTIVE : BOOL
END_METHOD

METHOD CALL_ERRORHANDLER
END_METHOD

METHOD CALL_ERRORHANDLER_STATECUTTING
END_METHOD

METHOD CALL_FBMETHODS
END_METHOD

METHOD CALL_FBMETHODS_BEFOREFLEXCAM
END_METHOD

METHOD CALL_FBMETHODS_CONTROLAXISBYPOS
END_METHOD

METHOD CALL_FB_CONTROLSETVALUES
END_METHOD

METHOD CALL_FB_DIFFERENTIATEPOSITION
END_METHOD

METHOD CALL_FM_CAMCREATOR_CONTINUOUS1
END_METHOD

METHOD CALL_FM_CAMCREATOR_CONTINUOUS2
END_METHOD

METHOD CALL_FM_CAMCREATOR_START
END_METHOD

METHOD CALL_FM_CAMCREATORS
END_METHOD

METHOD CALL_FM_FLEXCAM
END_METHOD

METHOD CALL_FM_FLEXCAM_INPUT
END_METHOD

METHOD CALL_INITDONE
END_METHOD

METHOD CALL_INITROUTINE
END_METHOD

METHOD CALL_INTERNALCTRL
END_METHOD

METHOD CALL_MASTEROFFSET
END_METHOD

METHOD CALL_MASTERTRIMM
END_METHOD

METHOD CALL_OUTPUT
END_METHOD

METHOD CALL_OUTPUTMINMAXVALUES
END_METHOD

METHOD CALL_OUTPUT_SF
END_METHOD

METHOD CALL_PARSYNCINCAM
END_METHOD

METHOD CALL_PARSYNCOUT
END_METHOD

METHOD CALL_REQUESTSSETCAMTABLE
END_METHOD

METHOD CALL_REQUESTSSETCAMTABLECTRL
END_METHOD

METHOD CALL_REQUESTS_EXT
END_METHOD

METHOD CALL_RESETCOMMANDS
END_METHOD

METHOD CALL_RESETOUTPUT
END_METHOD

METHOD CALL_RESETWARNINGS
END_METHOD

METHOD CALL_SETTOOLNOOUT
END_METHOD

METHOD CALL_STATEMACHINE
END_METHOD

METHOD CALL_ABC_INPUT_PROFILEPARAMETER
END_METHOD

METHOD CALL_CALCACTXKOORDINATEN
END_METHOD

METHOD CALL_CALCCAM_CONTINUOUS
END_METHOD

METHOD CALL_CALCCAM_START
END_METHOD

METHOD CALL_CALCSYNCARRAY
END_METHOD

METHOD CALL_CHECKCUTTINGPARCHANGES
END_METHOD

METHOD CALL_CONTINUOUSCAMSETYOFFSET
END_METHOD

METHOD CALL_CUTLENGTHCALCULATOR
END_METHOD

METHOD CALL_INIT_FLEXCAM
END_METHOD

METHOD CALL_LOCKCAMTABLE
END_METHOD

METHOD CALL_LOCKCROSSCUTTERPAR
END_METHOD

METHOD CALL_LOCKCUTTINGPAR
END_METHOD

METHOD CALL_LOCKCUTTINGPAR_ECCMODE_0
END_METHOD

METHOD CALL_LOCKCUTTINGPAR_ECCMODE_1
END_METHOD

METHOD CALL_PREPARENEXTCUT
END_METHOD

METHOD CALL_PREPARENEXTCUT_ECCMODEPAR
END_METHOD

METHOD CALL_RESETALLCAMCREATOR
END_METHOD

METHOD CALL_SEARCHACTYCOORDINATE
END_METHOD

METHOD CALL_SEARCHPARKPOS
END_METHOD

METHOD CALL_SETNEXTCAMCREATOR_CONTINUOUS
END_METHOD

METHOD CALL_YCOORDINATEMANAGER
END_METHOD

METHOD CHECKSLAVENOTINPARKPOS : BOOL
VAR_INPUT
	LRSETYPOS : LREAL;
	LRYSTART : LREAL;
	LRYPARK : LREAL;
	LRYEND : LREAL;
END_VAR
END_METHOD

METHOD CALL_CP_000_CYCLIC
END_METHOD

METHOD CALL_CP_001_INIT
END_METHOD

METHOD CALL_CP_001_INIT_OLD
END_METHOD

METHOD CALL_CP_141_IN_PARK_POS
END_METHOD

METHOD CALL_CP_142_ASYNC_PHASE
END_METHOD

METHOD CALL_CP_143_ENTRY_IN_SYNC_PHASE
END_METHOD

METHOD CALL_CP_143_ENTRY_IN_SYNC_PHASE_TRANSITION
END_METHOD

METHOD CALL_CP_144_EXIT_SYNC_PHASE
END_METHOD

METHOD CALL_CP_144_EXIT_SYNC_PHASE_TRANSITION
END_METHOD

METHOD CALL_CP_145_START_CAM
END_METHOD

METHOD CALL_CP_146_STOP_CAM
END_METHOD

METHOD CALL_CP_148_HOLD_IN_PARK_POS
END_METHOD

METHOD CALL_CP_148_HOLD_IN_PARK_POS_CONTINUECUTTING
END_METHOD

METHOD CALL_CP_148_HOLD_IN_PARK_POS_ENDOFPROFILE
END_METHOD

METHOD CALL_CP_802_STOP_IN_PARK_POS
END_METHOD

METHOD CALL_CP_900_DONE
END_METHOD

METHOD CALL_CUTTING_PROCESS
END_METHOD

METHOD CALL_S000_CYCLIC
END_METHOD

METHOD CALL_S002_STANDBY
END_METHOD

METHOD CALL_S030_SYNCHRONISING_POS
END_METHOD

METHOD CALL_S030_SYNCHRONISING_POS_ECCMODESELECT
END_METHOD

METHOD CALL_S030_SYNCHRONISING_POS_ECCMODE_0
END_METHOD

METHOD CALL_S030_SYNCHRONISING_POS_ECCMODE_1
END_METHOD

METHOD CALL_S032_POSITIONING_TO_START_POS
END_METHOD

METHOD CALL_S034_POSITIONING_TO_PARK_POS
END_METHOD

METHOD CALL_S035_CUTTING
END_METHOD

METHOD CALL_S996_STOP
END_METHOD

METHOD CALL_S999_ERROR
END_METHOD

METHOD CALL_T000_ALLSTATES
END_METHOD

METHOD CALL_S034_POSITIONING_TO_PARK_POS_OUT
END_METHOD

METHOD CALL_S035_CUTTING_OUT
END_METHOD

METHOD CALL_STATEMACHINE_OUT
END_METHOD

(* ---- L_TS2P_TM_CROSSCUTTERSTATE.fb ---- *)
FUNCTION_BLOCK L_TS2P_TM_CROSSCUTTERSTATE EXTENDS L_TS2P_TM_CrossCutterBase
VAR
	LRCYCMASTERPOS_INT : LREAL;
	XLOADREGPOS_INT : BOOL;
	LRLOADREGPOS_INT : LREAL;
	LRSETMOTORPRECTRLTRQOUT : LREAL;
	XREGISTERCTRLACTIVE : BOOL;
	XMARKRECEIVED_OLD : BOOL;
	XTEACHMARKWINDOW_OLD : BOOL;
	XLOADREGPOS_OLD : BOOL;
	_SCTPRECEIVEDATA : L_MC1P_TpReceiveData;
	_FB_TPRECDATAPROXYMARKCORR : L_MC1P_TouchProbeRecDataProxy;
	_FB_TPRECDATAPROXYTOOLCORR : L_MC1P_TouchProbeRecDataProxy;
	XMARKSENSORVALUESTORED_OLD : BOOL;
	AP11_XSETCUTLENGTHINPRODUCT_OLD : BOOL;
	EWARNINGID : WORD;
	FM_L_TS2P_MASTERVALUECORRECTION_LRACTVEL_OLD : LREAL;
	DNNUMAXISY_INT : DWORD := 1;
	DNDENAXISY_INT : DWORD := 1;
	XINVALIDCUTPRODUCTFORMAT : BOOL;
	XSCSCALINGVALID : BOOL := FALSE;
	XENABLETORQUEFOLLOWER : BOOL;
	XENABLEREGCTRLCORR : BOOL;
	XINVALIDTEACHMARKPOS : BOOL;
	XTPRECEIVED_INT : BOOL;
	LRTPACTPOSITION_INT : LREAL;
	XWARNINGINVALIDMARKRECIVED : BOOL;
	XTAKENEXTSTACKPOS : BOOL;
	LRSTACKLATESTDIST : LREAL;
	LRSENSORTOOLDIST_LOCK : LREAL;
	LRMARKPOS_LOCK : LREAL;
	XFIRSTCUTOFARRAY : BOOL;
	XCUTLENGTHINPRODUCTCHANGED_LOCK : BOOL;
	ISETNOCUTLENGTH_LOCK : INT;
	ISETNOOFMAXCUTLENGTH_LOCK : INT;
	LRUPPERCORRPOS_LOCK : LREAL;
	LRLOWERCORRPOS_LOCK : LREAL;
	ALRCUTLENGTHINPRODUCT_LOCK : ARRAY [1..10] OF LREAL;
	LRMARKSENSORPOS_LOCK : LREAL;
	LRREGISTERLENGTH_LOCK : LREAL;
	LRMINLOWERCORRPOS : LREAL;
	XCORRINSAMECYCLE : BOOL;
	LRFACTOR_NMOTOR_D_NAPPL : LREAL := 1;
	LRFACTOR_NAPPL_D_NMOTOR : LREAL := 1;
	LRFACTOR_MMOTOR_D_MAPPL : LREAL;
	INUMOFCUTLENGTH_LOCK : INT;
	INUMOFCUTLENGTH_INT : INT;
	LRREGPOS_ENDCUT : LREAL := 360;
	LRX_STOPCAMEND : LREAL := 360;
	_XSTACKENABLE : BOOL;
	_RC_LRUPPERCORRPOS : LREAL;
	_RC_LRLOWERCORRPOS : LREAL;
	_RC_XENABLE : BOOL;
	_RC_XMARKWINDOWOPEN : BOOL;
	_RC_XMARKOUTOFWINDOW : BOOL;
	_RC_XMARKNOTDETECTED : BOOL;
	_RC_XMARKWINDOWTEACHED : BOOL;
	_RC_LRGEARFACTORCORR : LREAL;
	_RC_XGEARFACTORCORRLIMITED : BOOL;
	_RC_LRPOSOUT : LREAL;
	_RC_LRACTVEL : LREAL;
	_RC_XERROR : BOOL;
	_RC_WERRORID : WORD;
	_RC_XLIMITACTIVE : BOOL;
	_RC_LRACTMARKERROR : LREAL;
	_RC_LRACTMARKDIST : LREAL;
	_RC_XINITDONE : BOOL;
	_RC_XCORRACTIVE : BOOL;
	_RC_XMARKRECEIVED : BOOL;
	_RC_LRREGMARKPOS : LREAL;
	_RC_XSETREGPOS2MASTERPOS : BOOL;
	LRACTMARKPOSDIFF : LREAL;
	FM_L_TS2P_MASTERVALUECORRECTION : L_TS2P_MasterValueCorrection;
	FM_L_TS2P_TOOLCORRECTION : L_TS2P_ToolCorrection;
	FB_L_TB2P_TP_CONVERTER : L_TB2P_TP_Converter;
	ITPCONVERTTPENABLECNTR : INT;
	FB_SETTORQUE1 : L_MC1P_SetTorqueOffset;
	FB_STACK : L_MB1P_Stack;
	WRESTART_LOCK : WORD;
	SCCAMTABLE_INT : MC_Cam_REF;
	SCSETXPROFILE_TEMP : L_MC2P_AxisProfile;
	SCSETYPROFILE_TEMP : L_MC2P_AxisProfile;
	PCAMDATA : POINTER TO L_MC2P_CamData;
	C_INUMOFCUTLENGTH : INT := 10;
END_VAR
END_FUNCTION_BLOCK

METHOD CALL_FM_TOOLCORRECTION : BOOL
END_METHOD

METHOD CALL_FM_TOOLCORRECTION_INPUT : BOOL
END_METHOD

METHOD CALL_ERRORHANDLER
END_METHOD

METHOD CALL_ERRORHANDLER_STATECUTTING
END_METHOD

METHOD CALL_FBMETHODS
END_METHOD

METHOD CALL_FBMETHODS_BEFOREFLEXCAM
END_METHOD

METHOD CALL_FBMETHODS_CONTROLAXISBYPOS
END_METHOD

METHOD CALL_FB_L_TB2P_TP_CONVERTER
END_METHOD

METHOD CALL_FB_SETTORQUE
END_METHOD

METHOD CALL_FB_SETTORQUE_INPUT
END_METHOD

METHOD CALL_FB_STACK
END_METHOD

METHOD CALL_FB_STACK_INPUT
END_METHOD

METHOD CALL_FM_CAMCREATOR_STANDSTILL
END_METHOD

METHOD CALL_FM_CAMCREATOR_STOP
END_METHOD

METHOD CALL_FM_CAMCREATORS
END_METHOD

METHOD CALL_FM_FLEXCAM
END_METHOD

METHOD CALL_FM_FLEXCAM_INPUT
END_METHOD

METHOD CALL_FM_REGISTERCONTROL
END_METHOD

METHOD CALL_FM_REGISTERCONTROL_INPUT
END_METHOD

METHOD CALL_FUN_GETSCALING
END_METHOD

METHOD CALL_INITDONE
END_METHOD

METHOD CALL_INITROUTINE
END_METHOD

METHOD CALL_INTERNALCTRL
END_METHOD

METHOD CALL_INTERNALCTRLBASEEXTENSION
END_METHOD

METHOD CALL_OUTPUT
END_METHOD

METHOD CALL_OUTPUTMINMAXVALUES
END_METHOD

METHOD CALL_OUTPUT_SF
END_METHOD

METHOD CALL_RESETCOMMANDS
END_METHOD

METHOD CALL_RESETOUTPUT
END_METHOD

METHOD CALL_RESETWARNINGS
END_METHOD

METHOD CALL_CALCCAM_RESTARTFROMSTOPCAM
END_METHOD

METHOD CALL_CALCCAM_STANDSTILL
END_METHOD

METHOD CALL_CALCCAM_STOP
END_METHOD

METHOD CALL_CALCSYNCARRAY_AP10STOPCAM
END_METHOD

METHOD CALL_CHECKARRAYOFCUTLENGTHCHANGES
END_METHOD

METHOD CALL_CHECKCUTPRODUCTFORMAT
END_METHOD

METHOD CALL_CHECKCUTTINGPARCHANGES
END_METHOD

METHOD CALL_CHECKRESTARTFROMSTOPCAM
END_METHOD

METHOD CALL_INIT_FLEXCAM
END_METHOD

METHOD CALL_LOCKCAMTABLE
END_METHOD

METHOD CALL_LOCKCROSSCUTTERPAR
END_METHOD

METHOD CALL_LOCKCUTTINGMODE
END_METHOD

METHOD CALL_LOCKCUTTINGPAR
END_METHOD

METHOD CALL_LOCKCUTTINGPAR_ECCMODE_2
END_METHOD

METHOD CALL_LOCKCUTTINGPAR_ECCMODE_3
END_METHOD

METHOD CALL_LOCKREGISTERCONTROLPAR
END_METHOD

METHOD CALL_PREAPAREARRAYOFCUTLENGTH
END_METHOD

METHOD CALL_PREPARENEXTCUT_ECCMODEPAR
END_METHOD

METHOD CALL_PREPARENEXTCUT_ECCMODEPAR_ECCMODE_2
END_METHOD

METHOD CALL_PREPARENEXTCUT_ECCMODEPAR_ECCMODE_3
END_METHOD

METHOD CALL_CP_000_CYCLIC
END_METHOD

METHOD CALL_CP_001_INIT
END_METHOD

METHOD CALL_CP_144_EXIT_SYNC_PHASE
END_METHOD

METHOD CALL_CP_148_HOLD_IN_PARK_POS
END_METHOD

METHOD CALL_CP_148_HOLD_IN_PARK_POS_CONTINUECUTTING
END_METHOD

METHOD CALL_CP_148_HOLD_IN_PARK_POS_ENDOFPROFILE
END_METHOD

METHOD CALL_CP_801_WAIT_OF_NEXT_CUT
END_METHOD

METHOD CALL_CP_802_STOP_IN_PARK_POS
END_METHOD

METHOD CALL_CP_900_DONE
END_METHOD

METHOD CALL_CUTTING_PROCESS
END_METHOD

METHOD CALL_S000_CYCLIC
END_METHOD

METHOD CALL_S002_READY
END_METHOD

METHOD CALL_S030_SYNCHRONISING_POS
END_METHOD

METHOD CALL_S030_SYNCHRONISING_POS_ECCMODESELECT
END_METHOD

METHOD CALL_S030_SYNCHRONISING_POS_ECCMODE_2
END_METHOD

METHOD CALL_S032_POSITIONING_TO_START_POS
END_METHOD

METHOD CALL_S999_ERROR
END_METHOD

(* ---- L_TS2P_TM_ELECTRONICGEARBOXBASE.fb ---- *)
FUNCTION_BLOCK L_TS2P_TM_ELECTRONICGEARBOXBASE EXTENDS L_TB2P_SyncMotionControl
VAR_OUTPUT
	PPAR : POINTER TO L_TS2P_scPar_TM_ElectronicGearboxBase;
	PSF : POINTER TO L_TS2P_scSF_TM_ElectronicGearboxBase;
	PAP : POINTER TO L_TS2P_scAP_TM_ElectronicGearboxBase;
END_VAR
VAR
	TM_ELECTRONICGEARBOXBASECONFIG : L_TB2P_ModuleHandlerConfig;
	PSCINPUT : POINTER TO L_TS2P_ElectronicGearboxBaseIn;
	PSCOUTPUT : POINTER TO L_TS2P_ElectronicGearboxBaseOut;
	XVELSYNCOUTTOBASESPEEDBUSY : BOOL;
	_LRSETBASEVEL : LREAL;
	XFM_SD_OFFSETBUSY : BOOL;
	_XSYNCHRONISEDBASEVEL : BOOL;
	XFM_SD_ACCDECBASEVEL : BOOL;
	_XSYNCOUTBASEVELDONE : BOOL;
	_XSYNCOUTBASEVELDONE_OLD : BOOL;
	_XSYNCOUTBASEVELDONE_RTRIG : BOOL;
	FM_L_TS2P_SYNCDRIVEVEL : L_TS2P_SyncDriveVel;
	XTRIMPOS_INT_OLD : BOOL;
	XTRIMNEG_INT_OLD : BOOL;
	_XSYNCVEL : BOOL;
	_XSYNCOUTINSTANT : BOOL;
	_LRVELOFFSET : LREAL;
	_LRPOSOFFSETTOTALPOS : LREAL;
	_LRPOSOFFSETTOTALVEL : LREAL;
	_LROFFSETTOTALVEL : LREAL;
	_LRSETTRIMOFFSETOUT : LREAL;
	_XSYNCOUTDONE : BOOL;
	_XSYNCOUTDONE_OLD : BOOL;
	_XSYNCOUTDONE_RTRIG : BOOL;
	_XSYNCHRONISED : BOOL;
	_XACCDECSYNC : BOOL;
	_XOFFSETTRIMBUSY : BOOL;
	DWGEARINGNUMERATOR_INT : DWORD;
	DWGEARINGDENOMINATOR_INT : DWORD;
	WMODE_INT : WORD;
	IACTMASTERDIRECTIONTMP : INT;
	XERROR_MODULOAXISISREQUIRED : BOOL;
	XERROR_INVALIDCOUPLINGMODE : BOOL;
	XWARNINGDIRECTIONDISABLEDSYNCINT : BOOL;
	XWARNINGDIRECTIONDISABLEDBASEVEL : BOOL;
	ETMSTATE_INT_TEMP : L_TB2P_States;
	XQSPAPPLICATION_OLD : BOOL;
	_XSYNCDRIVEENABLE : BOOL;
	_LRSYNCDRIVESETSLAVEVELOUT : LREAL;
	XENABLECONTROLSETVALUES : BOOL;
	FB_CONTROLSETVALUES : L_MC1P_ControlSetValues := STRUCT(eSetValueMode := L_MC1P_SetValueMode.VelAcc, xIgnoreAccForPosCalc := TRUE);
	FB_ALLOWEDDIRECTION : L_TS2P_AllowedDirection := STRUCT(eSetValueMode := L_MC1P_SetValueMode.VelAcc);
	XINVALIDBASEVELFLAG : BOOL;
	EERRORID_FIRST_OLD : L_IE1P_Error;
END_VAR
END_FUNCTION_BLOCK

METHOD CALL_FB_ALLOWEDDIRECTION
END_METHOD

METHOD CALL_ALLOCPOINTADR
END_METHOD

METHOD CALL_CTRLREQACTIVE : BOOL
END_METHOD

METHOD CALL_ERRORHANDLER
END_METHOD

METHOD CALL_FBMETHODS
END_METHOD

METHOD CALL_FB_CONTROLAXISBYVEL
END_METHOD

METHOD CALL_FB_CONTROLAXISBYVEL_INPUT
END_METHOD

METHOD CALL_FM_SYNCHRONIZEDDRIVE
END_METHOD

METHOD CALL_FM_SYNCHRONIZEDDRIVE_INPUT
END_METHOD

METHOD CALL_FM_SYNCHRONIZEDDRIVE_RESETFM
END_METHOD

METHOD CALL_INITDONE
END_METHOD

METHOD CALL_INITROUTINE
END_METHOD

METHOD CALL_INTERNALCTRL
END_METHOD

METHOD CALL_OUTPUT
END_METHOD

METHOD CALL_OUTPUT_SF
END_METHOD

METHOD CALL_REQUESTS_EXT
END_METHOD

METHOD CALL_RESETCOMMANDS
END_METHOD

METHOD CALL_RESETOUTPUT
END_METHOD

METHOD CALL_ABC_INPUT_PROFILEPARAMETER
END_METHOD

METHOD CALL_S000_CYCLIC
END_METHOD

METHOD CALL_S001_INIT
END_METHOD

METHOD CALL_S002_STANDBY
END_METHOD

METHOD CALL_S003_HOMING
END_METHOD

METHOD CALL_S010_JOGGING
END_METHOD

METHOD CALL_S030_ACC_DEC_SYNC
END_METHOD

METHOD CALL_S031_SYNCHRONISED
END_METHOD

METHOD CALL_S051_BASEVELOCITY
END_METHOD

METHOD CALL_S996_STOP
END_METHOD

METHOD CALL_S999_ERROR
END_METHOD

METHOD CALL_STATEMACHINE
END_METHOD

METHOD CALL_T000_ALLSTATES
END_METHOD

METHOD CALL_T030_ACC_DEC_SYNC
END_METHOD

METHOD CALL_T031_SYNCHRONISED
END_METHOD

METHOD CALL_T051_BASEVELOCITY
END_METHOD

METHOD CALL_050_ABORT
END_METHOD

METHOD CALL_S000_CYCLIC_OUT
END_METHOD

METHOD CALL_S003_HOMING_OUT
END_METHOD

METHOD CALL_S010_JOGGING_OUT
END_METHOD

METHOD CALL_S014_MOVEABS_OUT
END_METHOD

METHOD CALL_S015_MOVEREL_OUT
END_METHOD

METHOD CALL_S996_STOP_OUT
END_METHOD

METHOD CALL_S999_ERROR_OUT
END_METHOD

METHOD CALL_STATEMACHINE_OUT
END_METHOD

METHOD CALL_T000_ALLSTATES_OUT
END_METHOD

(* ---- L_TS2P_TM_FLEXCAM.fb ---- *)
FUNCTION_BLOCK L_TS2P_TM_FLEXCAM EXTENDS L_TB2M_TM_MotionControl
VAR
	TM_FLEXCAMHIGH : L_TB2P_ModuleHandlerConfig;
	HALT_FLEXCAM : INT := 16712;
	ITFFLEXCAMHIGH : L_TS2P_IFlexCam := THIS^;
	SCDATA_INT : L_TS2P_scData_TM_FlexCam;
	PDATA : POINTER TO L_TS2P_scData_TM_FlexCam := ADR(scData_Int);
	PPAR : POINTER TO L_TS2P_scPar_TM_FlexCam;
	PSF : POINTER TO L_TS2P_scSF_TM_FlexCam;
	PAP : POINTER TO L_TS2P_scAP_TM_FlexCam;
	PINPUT3 : POINTER TO L_TS2P_FlexCamHighIn;
	POUTPUT3 : POINTER TO L_TS2P_FlexCamHighOut;
	_ITFSTRUCTPROVIDERFLEXCAMHIGH : L_TS2P_IStructProviderFlexCamHigh;
	FB_CONDAXISMOVING : L_TB2P_AxisMoving;
	FB_CONDMASTERDIRECTION : L_TB2P_ConditionMasterDirection;
	FB_CONDLOCKTOCAM : L_TS2P_ConditionLockToCam;
	FB_CONDVALIDCAMTABLE : L_TS2P_ConditionValidCamTable;
	FB_CONDITIONLIMITERSYNCIN : L_TS2P_ConditionLimiterSyncIn;
	FB_CONDITIONCHECKHOMINGNEEDED : L_UBUP_ConditionInput;
	FB_CONDITIONJOGGINGACTIVE : L_UBUP_ConditionInput;
	FB_CONDCOLLECTCAMIN : L_UBUP_ConditionCollectionAND := STRUCT(aitfCondition := [fb_ConditionOperationEnabled, fb_ConditionLimiter, fb_CondLockToCam, fb_CondValidCamTable, fb_ConditionJoggingActive, fb_ConditionAxisNotStopping, fb_ConditionLimiterSyncIn, fb_ConditionCheckHomingNeeded]);
	FB_TRANSITION2LOCKTOCAM : L_UBUP_RequestTransitionLevel;
	FB_TRANSITION2MOVETOPARKPOSITION : L_UBUP_RequestTransitionEdge;
	FB_TRANSITION2CAMOUTHALT : L_UBUP_RequestTransitionEdge;
	FB_TRANSITION2CAMMING : L_UBUP_RequestTransitionLevel;
	FB_TRANSITION2FINDCLUTCHXPOS : L_UBUP_RequestTransitionEdge;
	WSETCAMTABLE_INT : WORD := 1;
	XSLAVEABSOLUTE_OLD : BOOL;
	XUPDATECURVE : BOOL;
	XCAMTABLEVALID_INT : BOOL;
	XCAMTABLEINTERNALVALID : BOOL;
	CAMTABLEINTERNAL : MC_CAM_REF;
	PCAMDATA : POINTER TO L_MC2P_CamData;
	_WFC_ENABLEMODE : WORD;
	_WFC_ENABLEMODE_OLD : WORD;
	_LRFC_SETXPOSOUT : LREAL;
	_LRFC_SETXVELOUT : LREAL;
	_LRFC_SETXACCOUT : LREAL;
	_LRFC_SETYPOSOUT : LREAL;
	_LRFC_SETYVELOUT : LREAL;
	_LRFC_SETYACCOUT : LREAL;
	_LRFC_OFFSETMASTER : LREAL;
	_LRFC_OFFSETSLAVE : LREAL;
	_XFC_CRITICALCYCLE : BOOL;
	_XFC_ENDOFPROFILE : BOOL;
	_XFC_ACCDECSYNC : BOOL;
	_XFC_CAMSYNCHRONISED : BOOL;
	_LRFC_SETSLAVEPOSOUT : LREAL;
	_LRFC_SETSLAVEVELOUT : LREAL;
	_LRFC_SETSLAVEACCOUT : LREAL;
	XCAMCHANGEINSTANT_OLD : BOOL;
	LRMASTERVEL_OLD : LREAL;
	LRMASTERVEL_OLD2 : LREAL;
	LRMASTERPOS_OLD : LREAL;
	XCONTROLSETVALUESBUSY_OLD : BOOL;
	XMASTERABSOLUTE_OLD : BOOL;
	XLOADCLUTCHPOS_OLD : BOOL;
	XCLUTCHCLOSEOLD : BOOL;
	LRENDOFPROFILEWINDOWSIZE : LREAL := 0;
	SCSETXPROFILE : L_MC2P_AxisProfile;
	SCSETYPROFILE : L_MC2P_AxisProfile;
	XERROR_INVALIDSYNCMODE : BOOL;
	XERROR_INVALIDCAMTABLE : BOOL;
	XWARNING_INVALIDCAMTABLE : BOOL;
	XCOMMUNICATION : BOOL;
	_MCS_CAMTABLEOUT : MC_CAM_REF;
	FB_CAMBASIC : L_MC2P_CamBasic;
	FB_CAMTABLEINFO1 : L_TS2P_CamTableInfo;
	FB_FINDCAMXVALUE : L_MC2A_FindCamXValue;
	FM_FLEXCAMSTATE1 : L_MC2P_FlexCamHigh := STRUCT(ePosCtrlDirection := L_MC2P_ReverseCtrlDirection.both);
	FB_MULTICAMSEQUENCER1 : L_TS2P_MultiCamSequencer;
	FB_CAMTABLEINFO2 : L_TS2P_CamTableInfo;
	FB_CAMTABLEINFO3 : L_TS2P_CamTableInfo;
	FB_CAMTABLEINFO4 : L_TS2P_CamTableInfo;
	FB_SYNCPOSRESTOREOFFSET : L_TS2P_OffsetAndTrim;
	FB_CLUTCHEXTENDEDBASE : L_TB2P_ClutchExtendedBase;
	FB_DIRECTION : L_TB2P_AllowedDirection;
	FB_SYNCIN : LockToMaster;
	ADDOFFSETCYCLIC : L_MC1P_AddOffsetCyclic;
	FB_ALLOWEDDIRECTION : L_TS2P_AllowedDirection;
	FB_CONTROLSETVALUES : L_MC1P_ControlSetValues;
	MASTERVALUES_INT : L_MC1P_SetAxisRefMasterValues;
	FB_MOVETOPARKPOS : MC_MoveAbsolute;
	FB_HALT : MC_Halt;
	FB_BLINKCLUTCH : L_USPP_Oscillator;
	FB_BLINKSYNCIN : L_USPP_Oscillator;
	XSYNCINOLD : BOOL;
	LRCYCLELENGTH : LREAL;
	ETRAVERSINGRANGE : L_MC1P_TraversingRange;
	XMASTERPARCHANGED : BOOL;
	_ITFREQUESTCONDITIONWARNINGHIGHPRIO : L_UBUP_IRequest;
	IVISFRAMESIGNALFLOW : INT;
	DIFRAMESF : DINT;
	CONNECTOR : __SYSTEM.IQueryInterface;
	FLEXCAMEXTENSION : L_TS2P_IFlexCam;
END_VAR
END_FUNCTION_BLOCK

METHOD CALL_CHECKCONSTANTVELOCITY
VAR_INPUT
	LRVELOCITYLASTCYCLE : LREAL;
END_VAR
VAR_OUTPUT
	XCONSTANTVELOCITY : BOOL;
END_VAR
END_METHOD

METHOD CALL_CURVESKETCHING
END_METHOD

METHOD CALL_FM_CAMTABLEINFO1
END_METHOD

METHOD CALL_FM_CAMTABLEINFO2
END_METHOD

METHOD CALL_FM_CAMTABLEINFO3
END_METHOD

METHOD CALL_FM_CAMTABLEINFO4
END_METHOD

METHOD CALL_OUTPUTMINMAXVALUES
END_METHOD

METHOD CALL_OUTPUTMINMAXVALUESMODULOOVERRUN
END_METHOD

METHOD CALL_OUTPUTMINMAXVALUESOFCAMTABLES1
END_METHOD

METHOD CALL_OUTPUTMINMAXVALUESOFCAMTABLES1_2_3_4
END_METHOD

METHOD GET_INTERNCAMTABLE : MC_CAM_REF
END_METHOD

METHOD GET_LRCAMXEND : LREAL
END_METHOD

METHOD GET_LRCAMXSTART : LREAL
END_METHOD

METHOD GET_LRCAMYEND : LREAL
END_METHOD

METHOD GET_LRCAMYSTART : LREAL
END_METHOD

METHOD GET_XCOMMUNICATION : BOOL
END_METHOD

METHOD HANDLEREJECTEDREQUEST : BOOL
VAR_INPUT
	ITFREQUESTANNOUNCED : L_UBUP_IRequest;
END_VAR
VAR_OUTPUT
	ITFALTERNATIVEREQUEST : L_UBUP_IRequest;
END_VAR
END_METHOD

METHOD CALLFBS
VAR_INPUT
	ECASE : L_UBUP_StateHandleCase;
END_VAR
END_METHOD

METHOD CALLSTATE
VAR_INPUT
	ITFSTATESERVER : L_UBUP_IStateServer;
	ISTATE : INT;
	ECASE : L_UBUP_StateHandleCase;
END_VAR
END_METHOD

METHOD CHECKTRANSITION
VAR_INPUT
	ITFSTATESERVER : L_UBUP_IStateServer;
END_VAR
END_METHOD

METHOD FINALIZECYCLE
END_METHOD

METHOD PREPARECYCLE
END_METHOD

METHOD SETADDMODULEINFO
VAR_INPUT
	ESUBCOMPTYPE : UDINT;
	SLICINFO : STRING(10);
END_VAR
END_METHOD

METHOD STIMULATETRANSITION
VAR_INPUT
	ECASE : L_UBUP_StateHandleCase;
END_VAR
END_METHOD

METHOD CALL_SETLOCALMASTERVALUES
END_METHOD

METHOD STATE_11_ACC_DEC_SYNC
VAR_INPUT
	ECASE : L_UBUP_StateHandleCase;
	ISTATESERVER : L_UBUP_IStateServer;
END_VAR
END_METHOD

METHOD STATE_12_MOVE_TO_PARKPOS
VAR_INPUT
	ECASE : L_UBUP_StateHandleCase;
	ISTATESERVER : L_UBUP_IStateServer;
END_VAR
END_METHOD

METHOD STATE_13_CAMMING
VAR_INPUT
	ECASE : L_UBUP_StateHandleCase;
	ISTATESERVER : L_UBUP_IStateServer;
END_VAR
END_METHOD

METHOD STATE_14_FIND_CLUTCH_X_POS
VAR_INPUT
	ECASE : L_UBUP_StateHandleCase;
	ISTATESERVER : L_UBUP_IStateServer;
END_VAR
END_METHOD

METHOD STATE_HALT_FLEXCAM
VAR_INPUT
	ECASE : L_UBUP_StateHandleCase;
	ITFSTATESERVER : L_UBUP_IStateServer;
END_VAR
END_METHOD

METHOD CAM
VAR_INPUT
	ITFTECHMODULE : L_TS2P_IFlexCam;
	XENABLE : BOOL;
	XSYNCCAM : BOOL;
	SCCAMTABLE : L_MC2P.MC_CAM_REF;
	LRCYCMASTERPOS : LREAL;
	LRCYCMASTERVEL : LREAL;
	LRCYCMASTERACC : LREAL;
	LRSLAVEPOS : LREAL;
	LRSLAVEVEL : LREAL;
	LRSLAVEACC : LREAL;
	EOFFSETMODEMASTER : L_TS2P_OffsetMode := L_TS2P_OffsetMode.x_zero;
	ESCALINGMODEMASTER : L_TS2P_ScalingMode := L_TS2P_ScalingMode.x_zero;
	EOFFSETMODESLAVE : L_TS2P_OffsetMode := L_TS2P_OffsetMode.x_zero;
	ESCALINGMODESLAVE : L_TS2P_ScalingMode := L_TS2P_ScalingMode.x_zero;
	LRSETOFFSETMASTER : LREAL;
	LRSETOFFSETSLAVE : LREAL;
	LRSETSCALINGMASTER : LREAL;
	LRSETSCALINGSLAVE : LREAL;
	LRPROFGENMASTERVEL : LREAL;
	LRPROFGENMASTERACC : LREAL;
	LRPROFGENMASTERDEC : LREAL;
	LRPROFGENMASTERJERK : LREAL;
	LRPROFGENSLAVEVEL : LREAL;
	LRPROFGENSLAVEACC : LREAL;
	LRPROFGENSLAVEDEC : LREAL;
	LRPROFGENSLAVEJERK : LREAL;
	XPERIODIC : BOOL;
	XCAMCHANGEINSTANT : BOOL;
	XMASTERABSOLUTE : BOOL;
	XSLAVEABSOLUTE : BOOL;
END_VAR
VAR_OUTPUT
	XERROR : BOOL;
	EERRORID : L_IE1P.L_IE1P_Error;
	LRSETPOSOUT : LREAL;
	LRSETVELOUT : LREAL;
	LRSETACCOUT : LREAL;
	LRSETXPOSOUT : LREAL;
	LRSETXVELOUT : LREAL;
	LRSETXACCOUT : LREAL;
	LRSETYPOSOUT : LREAL;
	LRSETYVELOUT : LREAL;
	LRSETYACCOUT : LREAL;
	XENDOFPROFILE : BOOL;
	LRSETOFFSETMASTEROUT : LREAL;
	LRSETOFFSETSLAVEOUT : LREAL;
	LRCONVERTMASTERTOXPOS : LREAL;
	LRCAMPROFILERPOSOUT : LREAL;
	LRCONVERTYTOSLAVEPOS : LREAL;
	XDONE : BOOL;
	XBUSY : BOOL;
END_VAR
END_METHOD

METHOD CAMSEQUENCER
VAR_INPUT
	ITFTECHMODULE : L_TS2P_IFlexCam;
	XENABLE : BOOL;
	XCAMSEQUENCER : BOOL;
	XENDOFPROFILEIN : BOOL;
	CAMTABLE1 : L_MC2P.MC_CAM_REF;
	CAMTABLE2 : L_MC2P.MC_CAM_REF;
	CAMTABLE3 : L_MC2P.MC_CAM_REF;
	CAMTABLE4 : L_MC2P.MC_CAM_REF;
	XCAMCHANGEINSTANT : BOOL;
	XLOADCAMTABLE : BOOL;
	WSETCAMTABLE : WORD;
	EMODE : L_TS2P_CamSequenceMode := L_TS2P_CamSequenceMode.CyclicCam1;
END_VAR
VAR_OUTPUT
	XERROR : BOOL;
	EERRORID : L_IE1P_Error;
	CAMTABLEOUT : L_MC2P.MC_CAM_REF;
	XCAMTABLEVALID : BOOL;
END_VAR
END_METHOD

METHOD CLUTCH
VAR_INPUT
	ITFTECHMODULE : L_TS2P_IFlexCam;
	XENABLE : BOOL;
	XCLUTCHCLOSE : BOOL;
	ECLUTCHINMODE : L_TS2P_ClutchInMode;
	ECLUTCHOUTMODE : L_TS2P_ClutchOutMode;
	EALLOWEDDIRECTION : L_TB2P_AllowedDirection;
	LRCLUTCHINDIST : LREAL;
	LRCLUTCHOUTDIST : LREAL;
	LRCLUTCHOUTPOSITION : LREAL;
	LRCYCLICMASTERPOS : LREAL;
	LRCYCLICMASTERVEL : LREAL;
	LRCYCLICMASTERACC : LREAL;
	LRCYCLICAXISPOS : LREAL;
	LRCYCLICAXISVEL : LREAL;
	LRCYCLICAXISACC : LREAL;
	ETRAVERSINGRANGE : L_MC1P_TraversingRange;
	LRCYCLELENGTH : LREAL;
END_VAR
VAR_OUTPUT
	XERROR : BOOL;
	EERRORID : L_IE1P.L_IE1P_Error;
	XBUSY : BOOL;
	XDONE : BOOL;
	XSYNCHRONISED : BOOL;
	XACCDECSYNC : BOOL;
	LRSETPOSOUT : LREAL;
	LRSETVELOUT : LREAL;
	LRSETACCOUT : LREAL;
END_VAR
END_METHOD

METHOD HALT : BOOL
VAR_INPUT
	ITFTECHMODULE : L_TS2P_IFlexCam;
	XEXECUTE : BOOL;
	LRDEC : LREAL := 100;
	LRJERK : LREAL := 0;
END_VAR
VAR_OUTPUT
	XBUSY : BOOL;
	XDONE : BOOL;
	XCOMMANDABORTED : BOOL;
END_VAR
VAR_IN_OUT
	AXIS : AXIS_REF;
END_VAR
END_METHOD

METHOD MOVETOPARKPOS : BOOL
VAR_INPUT
	ITFTECHMODULE : L_TS2P_IFlexCam;
	XEXECUTEMOVETOPARKPOS : BOOL;
	EMOVETOPARKPOSMODE : L_TS2P_CamStopMode;
	LRPARKPOSITION : LREAL := 180;
	EPOSITIONINGDIRECTION : L_TS2P_SyncDirection := L_TS2P_SyncDirection.PositiveDirection;
	LRPOSITIONINGVEL : LREAL := 10;
	LRPOSITIONINGACC : LREAL := 100;
	LRPOSITIONINGDEC : LREAL := 100;
	LRJERK : LREAL := 0;
END_VAR
VAR_OUTPUT
	XBUSY : BOOL;
	XDONE : BOOL;
	XCOMMANDABORTED : BOOL;
END_VAR
VAR_IN_OUT
	AXIS : AXIS_REF;
END_VAR
END_METHOD

METHOD POSITIONFOLLOWER
VAR_INPUT
	ITFTECHMODULE : L_TS2P_IFlexCam;
	XENABLE : BOOL;
	LRPOSITION : LREAL;
	LRVELOCITY : LREAL;
	LRACCELERATION : LREAL;
	ESETVALUEMODE : L_MC1P_SetValueMode;
END_VAR
VAR_OUTPUT
	XERROR : BOOL;
	EERRORID : L_IE1P.L_IE1P_Error;
	XBUSY : BOOL;
END_VAR
END_METHOD

METHOD SYNCIN
VAR_INPUT
	ITFTECHMODULE : L_TS2P_IFlexCam;
	XENABLE : BOOL;
	XSYNCIN : BOOL;
	XSYNCPOSRESTORE : BOOL;
	ESYNCMODE : L_TS2P_SyncInMode;
	ESYNCDIRECTION : L_TS2P_SyncDirection;
	LRSYNCVEL : LREAL;
	LRSYNCACC : LREAL;
	LRSYNCDEC : LREAL;
	LRSYNCJERK : LREAL;
	LRPARKPOSITION : LREAL;
	LRCYCLICMASTERPOS : LREAL;
	LRCYCLICMASTERVEL : LREAL;
	LRCYCLICMASTERACC : LREAL;
	LRCYCLICAXISPOS : LREAL;
	LRCYCLICAXISVEL : LREAL;
	LRCYCLICAXISACC : LREAL;
END_VAR
VAR_OUTPUT
	XERROR : BOOL;
	EERRORID : L_IE1P.L_IE1P_Error;
	XBUSY : BOOL;
	XDONE : BOOL;
	XSYNCHRONISED : BOOL;
	XACCDECSYNC : BOOL;
	LRSETPOSOUT : LREAL;
	LRSETVELOUT : LREAL;
	LRSETACCOUT : LREAL;
	LROFFSETSYNCPOS : LREAL;
END_VAR
VAR_IN_OUT
	AXIS : AXIS_REF;
END_VAR
END_METHOD

METHOD CALL_ALLOCPOINTADR
END_METHOD

METHOD CALL_EXIT_CALLFBS
END_METHOD

METHOD CALL_INIT_CALLFBS
END_METHOD

METHOD CALL_INTERNALCTRL
END_METHOD

METHOD CALL_RESETOUTPUT
END_METHOD

METHOD MAPTMSTATE
VAR_INPUT
	ETMSTATEINTERNAL : L_TB2P_States;
END_VAR
VAR_OUTPUT
	ETMSTATEEXTERNAL : L_TB2P_States;
END_VAR
END_METHOD

(* ---- L_TS2P_TM_FLEXCAMBASE.fb ---- *)
FUNCTION_BLOCK L_TS2P_TM_FLEXCAMBASE EXTENDS L_TB2P_SyncMotionControl
VAR_OUTPUT
	PAP : POINTER TO L_TS2P_scAP_TM_FlexCamState;
	PPAR : POINTER TO L_TS2P_scPar_TM_FlexCamState := ADR(scPar_int);
	PSF : POINTER TO L_TS2P_scSF_TM_FlexCamState;
END_VAR
VAR
	TM_FLEXCAMBASECONFIG : L_TB2P_ModuleHandlerConfig;
	PSCINPUT : POINTER TO L_TS2P_FlexCamStateIn;
	PSCOUTPUT : POINTER TO L_TS2P_FlexCamStateOut;
	SCPAR_INT : L_TS2P_scPar_TM_FlexCamState;
	XCAMMINGBUSY_INT : BOOL;
	XENABLECAMPROFILERSTANDBY_INT : BOOL := TRUE;
	XINTERNALCAMBASICACTIVE_INT : BOOL;
	XCAMCHANGEINSTANT_OLD : BOOL;
	LRMASTERVEL_OLD : LREAL;
	LRMASTERVEL_OLD2 : LREAL;
	LRMASTERPOS_OLD : LREAL;
	XCONTROLSETVALUESBUSY_OLD : BOOL;
	XMASTERABSOLUTE_OLD : BOOL;
	XCAMTABLEVALID_INT : BOOL;
	XERROR_INVALIDSYNCMODE : BOOL;
	XERROR_INVALIDCAMTABLE : BOOL;
	XWARNING_INVALIDCAMTABLE : BOOL;
	LRTRACEACCMAX_INT : LREAL;
	XCOMMUNICATION : BOOL;
	CAMTABLE_INIT : MC_CAM_REF;
	XMASTERPARCHANGED : BOOL;
	MASTERID : POINTER TO WORD;
	LRCYCLELENGTH : LREAL;
	ETRAVERSINGRANGE : LREAL;
	LRACTYPOS : LREAL;
	LRACTYVEL : LREAL;
	LRCAMYSTART : LREAL;
	LRCAMYEND : LREAL;
	LRACTIVESCALINGSLAVEINVERSE : LREAL;
	XCAMTABLEINTERNALVALID : BOOL;
	CAMTABLEINTERNAL : MC_CAM_REF;
	PCAMDATA : POINTER TO L_MC2P_CamData;
	_WFC_ENABLEMODE : WORD;
	_WFC_ENABLEMODE_OLD : WORD;
	_LRFC_SETXPOSOUT : LREAL;
	_LRFC_SETXVELOUT : LREAL;
	_LRFC_SETXACCOUT : LREAL;
	_LRFC_SETYPOSOUT : LREAL;
	_LRFC_SETYVELOUT : LREAL;
	_LRFC_SETYACCOUT : LREAL;
	_LRFC_OFFSETMASTER : LREAL;
	_LRFC_OFFSETSLAVE : LREAL;
	_XFC_CRITICALCYCLE : BOOL;
	_XFC_ENDOFPROFILE : BOOL;
	_XFC_ACCDECSYNC : BOOL;
	_XFC_CAMSYNCHRONISED : BOOL;
	_XFC_BUSY : BOOL;
	_XFC_DONE : BOOL;
	_XFC_ERROR : BOOL;
	_LRFC_SETSLAVEPOSOUT : LREAL;
	_LRFC_SETSLAVEVELOUT : LREAL;
	_LRFC_SETSLAVEACCOUT : LREAL;
	LRENDOFPROFILEWINDOWSIZE : LREAL := 0;
	MP_LRCONVERTMASTERTOXPOS : LREAL;
	MP_LRCAMPROFILERPOSOUT : LREAL;
	MP_LRCONVERTYTOSLAVEPOS : LREAL;
	MP_LWENDOFPROFILECHECKSUM : LWORD;
	MP_XENDOFPROFPOSITIVE : BOOL;
	MP_XENDOFPROFNEGATIVE : BOOL;
	SCSETXPROFILE : L_MC2P_AxisProfile;
	SCSETYPROFILE : L_MC2P_AxisProfile;
	FB_CAMBASIC : L_MC2P_CamBasic;
	FB_CONTROLSETVALUES : L_MC1P_ControlSetValues;
	FB_CAMTABLEINFO1 : L_TS2P_CamTableInfo;
END_VAR
END_FUNCTION_BLOCK

METHOD CALL_ALLOCPOINTADR
END_METHOD

METHOD CALL_AXISCONTROLBYPOS
END_METHOD

METHOD CALL_AXISCONTROLBYPOS_INPUT
END_METHOD

METHOD CALL_CAMBOUNDS
END_METHOD

METHOD CALL_CTRLREQACTIVE : BOOL
END_METHOD

METHOD CALL_CURVESKETCHING
END_METHOD

METHOD CALL_ERRORHANDLER
END_METHOD

METHOD CALL_FBMETHODS
END_METHOD

METHOD CALL_FB_CAMBASIC
END_METHOD

METHOD CALL_FM_CAMTABLEINFO1
END_METHOD

METHOD CALL_FM_FLEXCAM
END_METHOD

METHOD CALL_FM_FLEXCAM_INPUT
END_METHOD

METHOD CALL_INITDONE
END_METHOD

METHOD CALL_INITROUTINE
END_METHOD

METHOD CALL_INTERNALCTRL
END_METHOD

METHOD CALL_MASTERAXISREF
VAR_INPUT
	MASTERVALUES : L_MC1P_IAXIS_REF_MASTERVALUES;
END_VAR
END_METHOD

METHOD CALL_OUTPUT
END_METHOD

METHOD CALL_OUTPUTMINMAXVALUES
END_METHOD

METHOD CALL_OUTPUTMINMAXVALUESMODULOOVERRUN
END_METHOD

METHOD CALL_OUTPUTMINMAXVALUESOFCAMTABLES1
END_METHOD

METHOD CALL_OUTPUT_SF
END_METHOD

METHOD CALL_REQUESTS_EXT
END_METHOD

METHOD CALL_RESETCOMMANDS
END_METHOD

METHOD CALL_RESETOUTPUT
END_METHOD

METHOD CALL_STATEMACHINE
END_METHOD

METHOD CALL_ABC_INPUT_PROFILEPARAMETER
END_METHOD

METHOD CAMREFCHANGED : BOOL
VAR_IN_OUT
	CAMREFNEW : MC_CAM_REF;
	CAMREFOLD : MC_CAM_REF;
END_VAR
END_METHOD

METHOD CAMREFVALID : BOOL
VAR_INPUT
	CAMREF : MC_CAM_REF;
END_VAR
END_METHOD

METHOD GET_INTERNCAMTABLE : MC_CAM_REF
END_METHOD

METHOD GET_ECAMTYPE : L_MC2P_CamType
END_METHOD

METHOD GET_LRACTIVESCALINGSLAVE : LREAL
END_METHOD

METHOD GET_LRCAMXEND : LREAL
END_METHOD

METHOD GET_LRCAMXSTART : LREAL
END_METHOD

METHOD GET_LRCAMYEND : LREAL
END_METHOD

METHOD GET_LRCAMYSTART : LREAL
END_METHOD

METHOD GET_XCOMMUNICATION : BOOL
END_METHOD

METHOD RESET_SYSTEMFAULT
END_METHOD

METHOD SET_SYSTEMFAULT
VAR_INPUT
	IN : L_IE1P_Error;
END_VAR
END_METHOD

METHOD SET_ESTATE
VAR_INPUT
	IN : L_TB2P_States;
END_VAR
END_METHOD

METHOD CALL_S000_CYCLIC
END_METHOD

METHOD CALL_S002_STANDBY
END_METHOD

METHOD CALL_S112_CAMMING
END_METHOD

METHOD CALL_S112_CAMMING_RESTARTFLEXCAM
END_METHOD

METHOD CALL_S996_STOP
END_METHOD

METHOD CALL_S999_ERROR
END_METHOD

METHOD CALL_T000_ALLSTATES
END_METHOD

METHOD CALL_T002_STANDBY
END_METHOD

(* ---- L_TS2P_TM_FLEXCAMSTATE.fb ---- *)
FUNCTION_BLOCK L_TS2P_TM_FLEXCAMSTATE EXTENDS L_TS2P_TM_FlexCamBase
VAR
	XSLAVEABSOLUTE_OLD : BOOL;
	XUPDATECURVE : BOOL;
	_XMCS_ENABLE : BOOL;
	_MCS_CAMTABLEOUT : MC_CAM_REF;
	FM_FLEXCAMSTATE1 : L_MC2P_FlexCamHigh := STRUCT(ePosCtrlDirection := L_MC2P_ReverseCtrlDirection.both);
	FB_MULTICAMSEQUENCER1 : L_TS2P_MultiCamSequencer;
	FB_CAMTABLEINFO2 : L_TS2P_CamTableInfo;
	FB_CAMTABLEINFO3 : L_TS2P_CamTableInfo;
	FB_CAMTABLEINFO4 : L_TS2P_CamTableInfo;
END_VAR
END_FUNCTION_BLOCK

METHOD CALL_CURVESKETCHING
END_METHOD

METHOD CALL_ERRORHANDLER
END_METHOD

METHOD CALL_FBMETHODS
END_METHOD

METHOD CALL_FM_CAMTABLEINFO2
END_METHOD

METHOD CALL_FM_CAMTABLEINFO3
END_METHOD

METHOD CALL_FM_CAMTABLEINFO4
END_METHOD

METHOD CALL_FM_FLEXCAM
END_METHOD

METHOD CALL_FM_FLEXCAM_INPUT
END_METHOD

METHOD CALL_FM_MULTICAMSEQUENCER
END_METHOD

METHOD CALL_FM_MULTICAMSEQUENCER_INPUT
END_METHOD

METHOD CALL_FIRSTCYCLE
END_METHOD

METHOD CALL_INTERNALCTRL
END_METHOD

METHOD CALL_OUTPUT
END_METHOD

METHOD CALL_OUTPUTMINMAXVALUES
END_METHOD

METHOD CALL_OUTPUTMINMAXVALUESOFCAMTABLES1
END_METHOD

METHOD CALL_OUTPUTMINMAXVALUESOFCAMTABLES1_2_3_4
END_METHOD

METHOD CALL_OUTPUT_SF
END_METHOD

METHOD CALL_RESETCOMMANDS
END_METHOD

METHOD CALL_RESETCOMMANDSFLEXCAM
END_METHOD

METHOD CALL_RESETOUTPUT
END_METHOD

METHOD FUN_FMSYNCDIRCTION : L_MC2P_ClutchMode
VAR_INPUT
	ESYNCMODE : L_TS2P_SyncModeFlexCam;
END_VAR
END_METHOD

METHOD GET_INTERNCAMTABLE : MC_CAM_REF
END_METHOD

METHOD GET_LRACTIVESCALINGSLAVE : LREAL
END_METHOD

METHOD GET_LRCAMXEND : LREAL
END_METHOD

METHOD GET_LRCAMXSTART : LREAL
END_METHOD

METHOD GET_LRCAMYEND : LREAL
END_METHOD

METHOD GET_LRCAMYSTART : LREAL
END_METHOD

METHOD CALL_S112_CAMMING_RESTARTFLEXCAM
END_METHOD

(* ---- L_TS2P_TM_SYNCANDCORRECTIONSTATE.fb ---- *)
FUNCTION_BLOCK L_TS2P_TM_SYNCANDCORRECTIONSTATE EXTENDS L_TS2P_TM_SyncPosBase
VAR
	TM_SYNCANDCORRECTIONSTATECONFIG : L_TB2P_ModuleHandlerConfig;
	ITFSYNCANDCORRECTIONSTATE : L_TS2P_ISyncAndCorrectionState := THIS^;
	SCDATA_INTSC : L_TS2P_scData_TM_SyncAndCorrectionState;
	PAP_SC : POINTER TO L_TS2P_scAP_TM_SyncAndCorrectionState;
	PSF_SC : POINTER TO L_TS2P_scSF_TM_SyncAndCorrectionState;
	PDATASC : POINTER TO L_TS2P_scData_TM_SyncAndCorrectionState := ADR(scData_IntSC);
	PPAR_SC : POINTER TO L_TS2P_scPar_TM_SyncAndCorrectionState;
	PINPUT3 : POINTER TO L_TS2P_SyncAndCorrectionStateIn;
	POUTPUT3 : POINTER TO L_TS2P_SyncAndCorrectionStateOut;
	_ITFSTRUCTPROVIDERSYNCANDCORRECTION : L_TS2P_IStructProviderSyncAndCorrection;
	FM_L_TS2P_MASTERVALUECORRECTION : L_TS2P_MasterValueCorrection;
	FM_L_TS2P_TOOLCORRECTION : L_TS2P_ToolCorrection;
	FB_TPRECDATAPROXYMARKCORR : L_MC1P_TouchProbeRecDataProxy;
	FB_TPRECDATAPROXYTOOLCORR : L_MC1P_TouchProbeRecDataProxy;
	CONNECTOR : __SYSTEM.IQueryInterface;
	SYNCANDCORRECTIONSTATEEXTENSION : L_TS2P_ISyncAndCorrectionState;
	SYNCPOSBASEEXTENSION : L_TS2P_ISyncPosBase;
END_VAR
END_FUNCTION_BLOCK

METHOD CALLFBS
VAR_INPUT
	ECASE : L_UBUP_StateHandleCase;
END_VAR
END_METHOD

METHOD FINALIZECYCLE
END_METHOD

METHOD PREPARECYCLE
END_METHOD

METHOD SETADDMODULEINFO
VAR_INPUT
	ESUBCOMPTYPE : UDINT;
	SLICINFO : STRING(10);
END_VAR
END_METHOD

METHOD CALL_SETLOCALMASTERVALUES
END_METHOD

METHOD STATE_11_SYNC_ACC
VAR_INPUT
	ECASE : L_UBUP_StateHandleCase;
	ISTATESERVER : L_UBUP_IStateServer;
END_VAR
END_METHOD

METHOD CALL_FM_MASTERVALUECORRECTION
END_METHOD

METHOD CALL_FM_MASTERVALUECORRECTION_INPUT
END_METHOD

METHOD CALL_FM_TOOLCORRECTION : BOOL
END_METHOD

METHOD CALL_FM_TOOLCORRECTION_INPUT : BOOL
END_METHOD

METHOD CALL_ALLOCPOINTADR
END_METHOD

METHOD CALL_EXIT_CALLFBS
END_METHOD

METHOD CALL_INIT_CALLFBS
END_METHOD

METHOD CALL_INTERNALCTRL
END_METHOD

METHOD CALL_RESETOUTPUT
END_METHOD
